(* IEC 61131-3 sources: REFUSR/GP/Refusr.jl/samples (part 18) *)

(* ---- 5-MUX_vitae-roger-ships.st ---- *)
(*
This code implements a shuffled multiplexer with 5 control bits.
The control bits are: Data[N21], Data[N4], Data[N1], Data[N2], Data[N3]
The input bits are: Data[N7], Data[N8], Data[N5], Data[N20], Data[N23], Data[N24], Data[N9], Data[N25], Data[N22], Data[N6], Data[N10], Data[N26], Data[N14], Data[N11], Data[N29], Data[N15], Data[N12], Data[N13], Data[N19], Data[N16], Data[N17], Data[N18], Data[N32], Data[N27], Data[N30], Data[N33], Data[N31], Data[N34], Data[N35], Data[N28], Data[N36], Data[N37]

The symbolic expression is:
((((((((((((((((((((((((((((((((!(((((!(IN21)) & (!(IN4))) & (!(IN1))) & (!(IN2))) & (!(IN3)))) | IN7) & ((!((((IN21 & (!(IN4))) & (!(IN1))) & (!(IN2))) & (!(IN3)))) | IN8)) & ((!(((((!(IN21)) & IN4) & (!(IN1))) & (!(IN2))) & (!(IN3)))) | IN5)) & ((!((((IN21 & IN4) & (!(IN1))) & (!(IN2))) & (!(IN3)))) | IN20)) & ((!(((((!(IN21)) & (!(IN4))) & IN1) & (!(IN2))) & (!(IN3)))) | IN23)) & ((!((((IN21 & (!(IN4))) & IN1) & (!(IN2))) & (!(IN3)))) | IN24)) & ((!(((((!(IN21)) & IN4) & IN1) & (!(IN2))) & (!(IN3)))) | IN9)) & ((!((((IN21 & IN4) & IN1) & (!(IN2))) & (!(IN3)))) | IN25)) & ((!(((((!(IN21)) & (!(IN4))) & (!(IN1))) & IN2) & (!(IN3)))) | IN22)) & ((!((((IN21 & (!(IN4))) & (!(IN1))) & IN2) & (!(IN3)))) | IN6)) & ((!(((((!(IN21)) & IN4) & (!(IN1))) & IN2) & (!(IN3)))) | IN10)) & ((!((((IN21 & IN4) & (!(IN1))) & IN2) & (!(IN3)))) | IN26)) & ((!(((((!(IN21)) & (!(IN4))) & IN1) & IN2) & (!(IN3)))) | IN14)) & ((!((((IN21 & (!(IN4))) & IN1) & IN2) & (!(IN3)))) | IN11)) & ((!(((((!(IN21)) & IN4) & IN1) & IN2) & (!(IN3)))) | IN29)) & ((!((((IN21 & IN4) & IN1) & IN2) & (!(IN3)))) | IN15)) & ((!(((((!(IN21)) & (!(IN4))) & (!(IN1))) & (!(IN2))) & IN3)) | IN12)) & ((!((((IN21 & (!(IN4))) & (!(IN1))) & (!(IN2))) & IN3)) | IN13)) & ((!(((((!(IN21)) & IN4) & (!(IN1))) & (!(IN2))) & IN3)) | IN19)) & ((!((((IN21 & IN4) & (!(IN1))) & (!(IN2))) & IN3)) | IN16)) & ((!(((((!(IN21)) & (!(IN4))) & IN1) & (!(IN2))) & IN3)) | IN17)) & ((!((((IN21 & (!(IN4))) & IN1) & (!(IN2))) & IN3)) | IN18)) & ((!(((((!(IN21)) & IN4) & IN1) & (!(IN2))) & IN3)) | IN32)) & ((!((((IN21 & IN4) & IN1) & (!(IN2))) & IN3)) | IN27)) & ((!(((((!(IN21)) & (!(IN4))) & (!(IN1))) & IN2) & IN3)) | IN30)) & ((!((((IN21 & (!(IN4))) & (!(IN1))) & IN2) & IN3)) | IN33)) & ((!(((((!(IN21)) & IN4) & (!(IN1))) & IN2) & IN3)) | IN31)) & ((!((((IN21 & IN4) & (!(IN1))) & IN2) & IN3)) | IN34)) & ((!(((((!(IN21)) & (!(IN4))) & IN1) & IN2) & IN3)) | IN35)) & ((!((((IN21 & (!(IN4))) & IN1) & IN2) & IN3)) | IN28)) & ((!(((((!(IN21)) & IN4) & IN1) & IN2) & IN3)) | IN36)) & ((!((((IN21 & IN4) & IN1) & IN2) & IN3)) | IN37)

*)

FUNCTION_BLOCK F_CollectInput
  VAR_IN_OUT
      Data : ARRAY[1..40] OF BOOL;
  END_VAR
  VAR_INPUT
      TICK  : BOOL := 0;
      IN1   : BOOL := 0;
      IN2   : BOOL := 0;
      IN3   : BOOL := 0;
      IN4   : BOOL := 0;
      IN5   : BOOL := 0;
      RESET : BOOL := FALSE;
  END_VAR
  VAR_OUTPUT
      Finished : BOOL;
  END_VAR
  VAR
      j    : USINT := 1;
      tock : BOOL  := 0;
  END_VAR
  IF NOT RESET AND tock = NOT TICK THEN
      Data[j]   := IN1;
      Data[j+1] := IN2;
      Data[j+2] := IN3;
      Data[j+3] := IN4;
      Data[j+4] := IN5;
      j := j + 5;
      tock := TICK;
  ELSE
      j := 1;
      tock := 0;
  END_IF;
  Finished := (j > 40);
END_FUNCTION_BLOCK

PROGRAM Boiler
  VAR
    Data  : ARRAY[1..40] OF BOOL;
    Ready : BOOL;
    CollectInput : F_CollectInput;
  END_VAR
  VAR
    TICK     AT %IX1.0 : BOOL;
    IN1      AT %IX0.3 : BOOL;
    IN2      AT %IX0.4 : BOOL;
    IN3      AT %IX0.5 : BOOL;
    IN4      AT %IX0.6 : BOOL;
    IN5      AT %IX0.7 : BOOL;
    OutReady AT %QX0.0 : BOOL := FALSE;
    FeedNext AT %QX0.1 : BOOL := FALSE;
    Out      AT %QX0.2 : BOOL;
  END_VAR
  CollectInput(TICK:=TICK, IN1:=IN1, IN2:=IN2, IN3:=IN3, IN4:=IN4, IN5:=IN5);
  Ready := CollectInput.Finished;
  FeedNext := 1;
  IF Ready THEN
    Out := (((((((((((((((((((((((((((((((((NOT (((((NOT Data[21]) AND (NOT Data[4])) AND (NOT Data[1])) AND (NOT Data[2])) AND (NOT Data[3]))) OR Data[7]) AND ((NOT ((((Data[21] AND (NOT Data[4])) AND (NOT Data[1])) AND (NOT Data[2])) AND (NOT Data[3]))) OR Data[8])) AND ((NOT (((((NOT Data[21]) AND Data[4]) AND (NOT Data[1])) AND (NOT Data[2])) AND (NOT Data[3]))) OR Data[5])) AND ((NOT ((((Data[21] AND Data[4]) AND (NOT Data[1])) AND (NOT Data[2])) AND (NOT Data[3]))) OR Data[20])) AND ((NOT (((((NOT Data[21]) AND (NOT Data[4])) AND Data[1]) AND (NOT Data[2])) AND (NOT Data[3]))) OR Data[23])) AND ((NOT ((((Data[21] AND (NOT Data[4])) AND Data[1]) AND (NOT Data[2])) AND (NOT Data[3]))) OR Data[24])) AND ((NOT (((((NOT Data[21]) AND Data[4]) AND Data[1]) AND (NOT Data[2])) AND (NOT Data[3]))) OR Data[9])) AND ((NOT ((((Data[21] AND Data[4]) AND Data[1]) AND (NOT Data[2])) AND (NOT Data[3]))) OR Data[25])) AND ((NOT (((((NOT Data[21]) AND (NOT Data[4])) AND (NOT Data[1])) AND Data[2]) AND (NOT Data[3]))) OR Data[22])) AND ((NOT ((((Data[21] AND (NOT Data[4])) AND (NOT Data[1])) AND Data[2]) AND (NOT Data[3]))) OR Data[6])) AND ((NOT (((((NOT Data[21]) AND Data[4]) AND (NOT Data[1])) AND Data[2]) AND (NOT Data[3]))) OR Data[10])) AND ((NOT ((((Data[21] AND Data[4]) AND (NOT Data[1])) AND Data[2]) AND (NOT Data[3]))) OR Data[26])) AND ((NOT (((((NOT Data[21]) AND (NOT Data[4])) AND Data[1]) AND Data[2]) AND (NOT Data[3]))) OR Data[14])) AND ((NOT ((((Data[21] AND (NOT Data[4])) AND Data[1]) AND Data[2]) AND (NOT Data[3]))) OR Data[11])) AND ((NOT (((((NOT Data[21]) AND Data[4]) AND Data[1]) AND Data[2]) AND (NOT Data[3]))) OR Data[29])) AND ((NOT ((((Data[21] AND Data[4]) AND Data[1]) AND Data[2]) AND (NOT Data[3]))) OR Data[15])) AND ((NOT (((((NOT Data[21]) AND (NOT Data[4])) AND (NOT Data[1])) AND (NOT Data[2])) AND Data[3])) OR Data[12])) AND ((NOT ((((Data[21] AND (NOT Data[4])) AND (NOT Data[1])) AND (NOT Data[2])) AND Data[3])) OR Data[13])) AND ((NOT (((((NOT Data[21]) AND Data[4]) AND (NOT Data[1])) AND (NOT Data[2])) AND Data[3])) OR Data[19])) AND ((NOT ((((Data[21] AND Data[4]) AND (NOT Data[1])) AND (NOT Data[2])) AND Data[3])) OR Data[16])) AND ((NOT (((((NOT Data[21]) AND (NOT Data[4])) AND Data[1]) AND (NOT Data[2])) AND Data[3])) OR Data[17])) AND ((NOT ((((Data[21] AND (NOT Data[4])) AND Data[1]) AND (NOT Data[2])) AND Data[3])) OR Data[18])) AND ((NOT (((((NOT Data[21]) AND Data[4]) AND Data[1]) AND (NOT Data[2])) AND Data[3])) OR Data[32])) AND ((NOT ((((Data[21] AND Data[4]) AND Data[1]) AND (NOT Data[2])) AND Data[3])) OR Data[27])) AND ((NOT (((((NOT Data[21]) AND (NOT Data[4])) AND (NOT Data[1])) AND Data[2]) AND Data[3])) OR Data[30])) AND ((NOT ((((Data[21] AND (NOT Data[4])) AND (NOT Data[1])) AND Data[2]) AND Data[3])) OR Data[33])) AND ((NOT (((((NOT Data[21]) AND Data[4]) AND (NOT Data[1])) AND Data[2]) AND Data[3])) OR Data[31])) AND ((NOT ((((Data[21] AND Data[4]) AND (NOT Data[1])) AND Data[2]) AND Data[3])) OR Data[34])) AND ((NOT (((((NOT Data[21]) AND (NOT Data[4])) AND Data[1]) AND Data[2]) AND Data[3])) OR Data[35])) AND ((NOT ((((Data[21] AND (NOT Data[4])) AND Data[1]) AND Data[2]) AND Data[3])) OR Data[28])) AND ((NOT (((((NOT Data[21]) AND Data[4]) AND Data[1]) AND Data[2]) AND Data[3])) OR Data[36])) AND ((NOT ((((Data[21] AND Data[4]) AND Data[1]) AND Data[2]) AND Data[3])) OR Data[37]));
    OutReady := 1;
    CollectInput(RESET:=TRUE);
  END_IF;
END_PROGRAM

CONFIGURATION Config0
  RESOURCE Res0 ON PLC
    TASK task0(INTERVAL := T#20ms,PRIORITY := 0);
    PROGRAM instance0 WITH task0 : Boiler;
  END_RESOURCE
END_CONFIGURATION

(* ---- 5-MUX_vodka-chive-wrier.st ---- *)
(*
This code implements a shuffled multiplexer with 5 control bits.
The control bits are: Data[N2], Data[N1], Data[N23], Data[N3], Data[N20]
The input bits are: Data[N6], Data[N11], Data[N7], Data[N5], Data[N22], Data[N21], Data[N24], Data[N25], Data[N8], Data[N4], Data[N9], Data[N10], Data[N12], Data[N13], Data[N26], Data[N27], Data[N28], Data[N15], Data[N29], Data[N14], Data[N18], Data[N34], Data[N31], Data[N16], Data[N17], Data[N19], Data[N35], Data[N32], Data[N30], Data[N37], Data[N36], Data[N33]

The symbolic expression is:
((((((((((((((((((((((((((((((((!(((((!(IN2)) & (!(IN1))) & (!(IN23))) & (!(IN3))) & (!(IN20)))) | IN6) & ((!((((IN2 & (!(IN1))) & (!(IN23))) & (!(IN3))) & (!(IN20)))) | IN11)) & ((!(((((!(IN2)) & IN1) & (!(IN23))) & (!(IN3))) & (!(IN20)))) | IN7)) & ((!((((IN2 & IN1) & (!(IN23))) & (!(IN3))) & (!(IN20)))) | IN5)) & ((!(((((!(IN2)) & (!(IN1))) & IN23) & (!(IN3))) & (!(IN20)))) | IN22)) & ((!((((IN2 & (!(IN1))) & IN23) & (!(IN3))) & (!(IN20)))) | IN21)) & ((!(((((!(IN2)) & IN1) & IN23) & (!(IN3))) & (!(IN20)))) | IN24)) & ((!((((IN2 & IN1) & IN23) & (!(IN3))) & (!(IN20)))) | IN25)) & ((!(((((!(IN2)) & (!(IN1))) & (!(IN23))) & IN3) & (!(IN20)))) | IN8)) & ((!((((IN2 & (!(IN1))) & (!(IN23))) & IN3) & (!(IN20)))) | IN4)) & ((!(((((!(IN2)) & IN1) & (!(IN23))) & IN3) & (!(IN20)))) | IN9)) & ((!((((IN2 & IN1) & (!(IN23))) & IN3) & (!(IN20)))) | IN10)) & ((!(((((!(IN2)) & (!(IN1))) & IN23) & IN3) & (!(IN20)))) | IN12)) & ((!((((IN2 & (!(IN1))) & IN23) & IN3) & (!(IN20)))) | IN13)) & ((!(((((!(IN2)) & IN1) & IN23) & IN3) & (!(IN20)))) | IN26)) & ((!((((IN2 & IN1) & IN23) & IN3) & (!(IN20)))) | IN27)) & ((!(((((!(IN2)) & (!(IN1))) & (!(IN23))) & (!(IN3))) & IN20)) | IN28)) & ((!((((IN2 & (!(IN1))) & (!(IN23))) & (!(IN3))) & IN20)) | IN15)) & ((!(((((!(IN2)) & IN1) & (!(IN23))) & (!(IN3))) & IN20)) | IN29)) & ((!((((IN2 & IN1) & (!(IN23))) & (!(IN3))) & IN20)) | IN14)) & ((!(((((!(IN2)) & (!(IN1))) & IN23) & (!(IN3))) & IN20)) | IN18)) & ((!((((IN2 & (!(IN1))) & IN23) & (!(IN3))) & IN20)) | IN34)) & ((!(((((!(IN2)) & IN1) & IN23) & (!(IN3))) & IN20)) | IN31)) & ((!((((IN2 & IN1) & IN23) & (!(IN3))) & IN20)) | IN16)) & ((!(((((!(IN2)) & (!(IN1))) & (!(IN23))) & IN3) & IN20)) | IN17)) & ((!((((IN2 & (!(IN1))) & (!(IN23))) & IN3) & IN20)) | IN19)) & ((!(((((!(IN2)) & IN1) & (!(IN23))) & IN3) & IN20)) | IN35)) & ((!((((IN2 & IN1) & (!(IN23))) & IN3) & IN20)) | IN32)) & ((!(((((!(IN2)) & (!(IN1))) & IN23) & IN3) & IN20)) | IN30)) & ((!((((IN2 & (!(IN1))) & IN23) & IN3) & IN20)) | IN37)) & ((!(((((!(IN2)) & IN1) & IN23) & IN3) & IN20)) | IN36)) & ((!((((IN2 & IN1) & IN23) & IN3) & IN20)) | IN33)

*)

FUNCTION_BLOCK F_CollectInput
  VAR_IN_OUT
      Data : ARRAY[1..40] OF BOOL;
  END_VAR
  VAR_INPUT
      TICK  : BOOL := 0;
      IN1   : BOOL := 0;
      IN2   : BOOL := 0;
      IN3   : BOOL := 0;
      IN4   : BOOL := 0;
      IN5   : BOOL := 0;
      RESET : BOOL := FALSE;
  END_VAR
  VAR_OUTPUT
      Finished : BOOL;
  END_VAR
  VAR
      j    : USINT := 1;
      tock : BOOL  := 0;
  END_VAR
  IF NOT RESET AND tock = NOT TICK THEN
      Data[j]   := IN1;
      Data[j+1] := IN2;
      Data[j+2] := IN3;
      Data[j+3] := IN4;
      Data[j+4] := IN5;
      j := j + 5;
      tock := TICK;
  ELSE
      j := 1;
      tock := 0;
  END_IF;
  Finished := (j > 40);
END_FUNCTION_BLOCK

PROGRAM Boiler
  VAR
    Data  : ARRAY[1..40] OF BOOL;
    Ready : BOOL;
    CollectInput : F_CollectInput;
  END_VAR
  VAR
    TICK     AT %IX1.0 : BOOL;
    IN1      AT %IX0.3 : BOOL;
    IN2      AT %IX0.4 : BOOL;
    IN3      AT %IX0.5 : BOOL;
    IN4      AT %IX0.6 : BOOL;
    IN5      AT %IX0.7 : BOOL;
    OutReady AT %QX0.0 : BOOL := FALSE;
    FeedNext AT %QX0.1 : BOOL := FALSE;
    Out      AT %QX0.2 : BOOL;
  END_VAR
  CollectInput(TICK:=TICK, IN1:=IN1, IN2:=IN2, IN3:=IN3, IN4:=IN4, IN5:=IN5);
  Ready := CollectInput.Finished;
  FeedNext := 1;
  IF Ready THEN
    Out := (((((((((((((((((((((((((((((((((NOT (((((NOT Data[2]) AND (NOT Data[1])) AND (NOT Data[23])) AND (NOT Data[3])) AND (NOT Data[20]))) OR Data[6]) AND ((NOT ((((Data[2] AND (NOT Data[1])) AND (NOT Data[23])) AND (NOT Data[3])) AND (NOT Data[20]))) OR Data[11])) AND ((NOT (((((NOT Data[2]) AND Data[1]) AND (NOT Data[23])) AND (NOT Data[3])) AND (NOT Data[20]))) OR Data[7])) AND ((NOT ((((Data[2] AND Data[1]) AND (NOT Data[23])) AND (NOT Data[3])) AND (NOT Data[20]))) OR Data[5])) AND ((NOT (((((NOT Data[2]) AND (NOT Data[1])) AND Data[23]) AND (NOT Data[3])) AND (NOT Data[20]))) OR Data[22])) AND ((NOT ((((Data[2] AND (NOT Data[1])) AND Data[23]) AND (NOT Data[3])) AND (NOT Data[20]))) OR Data[21])) AND ((NOT (((((NOT Data[2]) AND Data[1]) AND Data[23]) AND (NOT Data[3])) AND (NOT Data[20]))) OR Data[24])) AND ((NOT ((((Data[2] AND Data[1]) AND Data[23]) AND (NOT Data[3])) AND (NOT Data[20]))) OR Data[25])) AND ((NOT (((((NOT Data[2]) AND (NOT Data[1])) AND (NOT Data[23])) AND Data[3]) AND (NOT Data[20]))) OR Data[8])) AND ((NOT ((((Data[2] AND (NOT Data[1])) AND (NOT Data[23])) AND Data[3]) AND (NOT Data[20]))) OR Data[4])) AND ((NOT (((((NOT Data[2]) AND Data[1]) AND (NOT Data[23])) AND Data[3]) AND (NOT Data[20]))) OR Data[9])) AND ((NOT ((((Data[2] AND Data[1]) AND (NOT Data[23])) AND Data[3]) AND (NOT Data[20]))) OR Data[10])) AND ((NOT (((((NOT Data[2]) AND (NOT Data[1])) AND Data[23]) AND Data[3]) AND (NOT Data[20]))) OR Data[12])) AND ((NOT ((((Data[2] AND (NOT Data[1])) AND Data[23]) AND Data[3]) AND (NOT Data[20]))) OR Data[13])) AND ((NOT (((((NOT Data[2]) AND Data[1]) AND Data[23]) AND Data[3]) AND (NOT Data[20]))) OR Data[26])) AND ((NOT ((((Data[2] AND Data[1]) AND Data[23]) AND Data[3]) AND (NOT Data[20]))) OR Data[27])) AND ((NOT (((((NOT Data[2]) AND (NOT Data[1])) AND (NOT Data[23])) AND (NOT Data[3])) AND Data[20])) OR Data[28])) AND ((NOT ((((Data[2] AND (NOT Data[1])) AND (NOT Data[23])) AND (NOT Data[3])) AND Data[20])) OR Data[15])) AND ((NOT (((((NOT Data[2]) AND Data[1]) AND (NOT Data[23])) AND (NOT Data[3])) AND Data[20])) OR Data[29])) AND ((NOT ((((Data[2] AND Data[1]) AND (NOT Data[23])) AND (NOT Data[3])) AND Data[20])) OR Data[14])) AND ((NOT (((((NOT Data[2]) AND (NOT Data[1])) AND Data[23]) AND (NOT Data[3])) AND Data[20])) OR Data[18])) AND ((NOT ((((Data[2] AND (NOT Data[1])) AND Data[23]) AND (NOT Data[3])) AND Data[20])) OR Data[34])) AND ((NOT (((((NOT Data[2]) AND Data[1]) AND Data[23]) AND (NOT Data[3])) AND Data[20])) OR Data[31])) AND ((NOT ((((Data[2] AND Data[1]) AND Data[23]) AND (NOT Data[3])) AND Data[20])) OR Data[16])) AND ((NOT (((((NOT Data[2]) AND (NOT Data[1])) AND (NOT Data[23])) AND Data[3]) AND Data[20])) OR Data[17])) AND ((NOT ((((Data[2] AND (NOT Data[1])) AND (NOT Data[23])) AND Data[3]) AND Data[20])) OR Data[19])) AND ((NOT (((((NOT Data[2]) AND Data[1]) AND (NOT Data[23])) AND Data[3]) AND Data[20])) OR Data[35])) AND ((NOT ((((Data[2] AND Data[1]) AND (NOT Data[23])) AND Data[3]) AND Data[20])) OR Data[32])) AND ((NOT (((((NOT Data[2]) AND (NOT Data[1])) AND Data[23]) AND Data[3]) AND Data[20])) OR Data[30])) AND ((NOT ((((Data[2] AND (NOT Data[1])) AND Data[23]) AND Data[3]) AND Data[20])) OR Data[37])) AND ((NOT (((((NOT Data[2]) AND Data[1]) AND Data[23]) AND Data[3]) AND Data[20])) OR Data[36])) AND ((NOT ((((Data[2] AND Data[1]) AND Data[23]) AND Data[3]) AND Data[20])) OR Data[33]));
    OutReady := 1;
    CollectInput(RESET:=TRUE);
  END_IF;
END_PROGRAM

CONFIGURATION Config0
  RESOURCE Res0 ON PLC
    TASK task0(INTERVAL := T#20ms,PRIORITY := 0);
    PROGRAM instance0 WITH task0 : Boiler;
  END_RESOURCE
END_CONFIGURATION

(* ---- 5-MUX_wager-river-honky.st ---- *)
(*
This code implements a shuffled multiplexer with 5 control bits.
The control bits are: Data[N22], Data[N21], Data[N2], Data[N20], Data[N5]
The input bits are: Data[N3], Data[N6], Data[N4], Data[N8], Data[N23], Data[N9], Data[N7], Data[N24], Data[N25], Data[N1], Data[N14], Data[N26], Data[N28], Data[N15], Data[N13], Data[N27], Data[N10], Data[N29], Data[N17], Data[N33], Data[N11], Data[N12], Data[N16], Data[N30], Data[N19], Data[N18], Data[N31], Data[N36], Data[N37], Data[N34], Data[N32], Data[N35]

The symbolic expression is:
((((((((((((((((((((((((((((((((!(((((!(IN22)) & (!(IN21))) & (!(IN2))) & (!(IN20))) & (!(IN5)))) | IN3) & ((!((((IN22 & (!(IN21))) & (!(IN2))) & (!(IN20))) & (!(IN5)))) | IN6)) & ((!(((((!(IN22)) & IN21) & (!(IN2))) & (!(IN20))) & (!(IN5)))) | IN4)) & ((!((((IN22 & IN21) & (!(IN2))) & (!(IN20))) & (!(IN5)))) | IN8)) & ((!(((((!(IN22)) & (!(IN21))) & IN2) & (!(IN20))) & (!(IN5)))) | IN23)) & ((!((((IN22 & (!(IN21))) & IN2) & (!(IN20))) & (!(IN5)))) | IN9)) & ((!(((((!(IN22)) & IN21) & IN2) & (!(IN20))) & (!(IN5)))) | IN7)) & ((!((((IN22 & IN21) & IN2) & (!(IN20))) & (!(IN5)))) | IN24)) & ((!(((((!(IN22)) & (!(IN21))) & (!(IN2))) & IN20) & (!(IN5)))) | IN25)) & ((!((((IN22 & (!(IN21))) & (!(IN2))) & IN20) & (!(IN5)))) | IN1)) & ((!(((((!(IN22)) & IN21) & (!(IN2))) & IN20) & (!(IN5)))) | IN14)) & ((!((((IN22 & IN21) & (!(IN2))) & IN20) & (!(IN5)))) | IN26)) & ((!(((((!(IN22)) & (!(IN21))) & IN2) & IN20) & (!(IN5)))) | IN28)) & ((!((((IN22 & (!(IN21))) & IN2) & IN20) & (!(IN5)))) | IN15)) & ((!(((((!(IN22)) & IN21) & IN2) & IN20) & (!(IN5)))) | IN13)) & ((!((((IN22 & IN21) & IN2) & IN20) & (!(IN5)))) | IN27)) & ((!(((((!(IN22)) & (!(IN21))) & (!(IN2))) & (!(IN20))) & IN5)) | IN10)) & ((!((((IN22 & (!(IN21))) & (!(IN2))) & (!(IN20))) & IN5)) | IN29)) & ((!(((((!(IN22)) & IN21) & (!(IN2))) & (!(IN20))) & IN5)) | IN17)) & ((!((((IN22 & IN21) & (!(IN2))) & (!(IN20))) & IN5)) | IN33)) & ((!(((((!(IN22)) & (!(IN21))) & IN2) & (!(IN20))) & IN5)) | IN11)) & ((!((((IN22 & (!(IN21))) & IN2) & (!(IN20))) & IN5)) | IN12)) & ((!(((((!(IN22)) & IN21) & IN2) & (!(IN20))) & IN5)) | IN16)) & ((!((((IN22 & IN21) & IN2) & (!(IN20))) & IN5)) | IN30)) & ((!(((((!(IN22)) & (!(IN21))) & (!(IN2))) & IN20) & IN5)) | IN19)) & ((!((((IN22 & (!(IN21))) & (!(IN2))) & IN20) & IN5)) | IN18)) & ((!(((((!(IN22)) & IN21) & (!(IN2))) & IN20) & IN5)) | IN31)) & ((!((((IN22 & IN21) & (!(IN2))) & IN20) & IN5)) | IN36)) & ((!(((((!(IN22)) & (!(IN21))) & IN2) & IN20) & IN5)) | IN37)) & ((!((((IN22 & (!(IN21))) & IN2) & IN20) & IN5)) | IN34)) & ((!(((((!(IN22)) & IN21) & IN2) & IN20) & IN5)) | IN32)) & ((!((((IN22 & IN21) & IN2) & IN20) & IN5)) | IN35)

*)

FUNCTION_BLOCK F_CollectInput
  VAR_IN_OUT
      Data : ARRAY[1..40] OF BOOL;
  END_VAR
  VAR_INPUT
      TICK  : BOOL := 0;
      IN1   : BOOL := 0;
      IN2   : BOOL := 0;
      IN3   : BOOL := 0;
      IN4   : BOOL := 0;
      IN5   : BOOL := 0;
      RESET : BOOL := FALSE;
  END_VAR
  VAR_OUTPUT
      Finished : BOOL;
  END_VAR
  VAR
      j    : USINT := 1;
      tock : BOOL  := 0;
  END_VAR
  IF NOT RESET AND tock = NOT TICK THEN
      Data[j]   := IN1;
      Data[j+1] := IN2;
      Data[j+2] := IN3;
      Data[j+3] := IN4;
      Data[j+4] := IN5;
      j := j + 5;
      tock := TICK;
  ELSE
      j := 1;
      tock := 0;
  END_IF;
  Finished := (j > 40);
END_FUNCTION_BLOCK

PROGRAM Boiler
  VAR
    Data  : ARRAY[1..40] OF BOOL;
    Ready : BOOL;
    CollectInput : F_CollectInput;
  END_VAR
  VAR
    TICK     AT %IX1.0 : BOOL;
    IN1      AT %IX0.3 : BOOL;
    IN2      AT %IX0.4 : BOOL;
    IN3      AT %IX0.5 : BOOL;
    IN4      AT %IX0.6 : BOOL;
    IN5      AT %IX0.7 : BOOL;
    OutReady AT %QX0.0 : BOOL := FALSE;
    FeedNext AT %QX0.1 : BOOL := FALSE;
    Out      AT %QX0.2 : BOOL;
  END_VAR
  CollectInput(TICK:=TICK, IN1:=IN1, IN2:=IN2, IN3:=IN3, IN4:=IN4, IN5:=IN5);
  Ready := CollectInput.Finished;
  FeedNext := 1;
  IF Ready THEN
    Out := (((((((((((((((((((((((((((((((((NOT (((((NOT Data[22]) AND (NOT Data[21])) AND (NOT Data[2])) AND (NOT Data[20])) AND (NOT Data[5]))) OR Data[3]) AND ((NOT ((((Data[22] AND (NOT Data[21])) AND (NOT Data[2])) AND (NOT Data[20])) AND (NOT Data[5]))) OR Data[6])) AND ((NOT (((((NOT Data[22]) AND Data[21]) AND (NOT Data[2])) AND (NOT Data[20])) AND (NOT Data[5]))) OR Data[4])) AND ((NOT ((((Data[22] AND Data[21]) AND (NOT Data[2])) AND (NOT Data[20])) AND (NOT Data[5]))) OR Data[8])) AND ((NOT (((((NOT Data[22]) AND (NOT Data[21])) AND Data[2]) AND (NOT Data[20])) AND (NOT Data[5]))) OR Data[23])) AND ((NOT ((((Data[22] AND (NOT Data[21])) AND Data[2]) AND (NOT Data[20])) AND (NOT Data[5]))) OR Data[9])) AND ((NOT (((((NOT Data[22]) AND Data[21]) AND Data[2]) AND (NOT Data[20])) AND (NOT Data[5]))) OR Data[7])) AND ((NOT ((((Data[22] AND Data[21]) AND Data[2]) AND (NOT Data[20])) AND (NOT Data[5]))) OR Data[24])) AND ((NOT (((((NOT Data[22]) AND (NOT Data[21])) AND (NOT Data[2])) AND Data[20]) AND (NOT Data[5]))) OR Data[25])) AND ((NOT ((((Data[22] AND (NOT Data[21])) AND (NOT Data[2])) AND Data[20]) AND (NOT Data[5]))) OR Data[1])) AND ((NOT (((((NOT Data[22]) AND Data[21]) AND (NOT Data[2])) AND Data[20]) AND (NOT Data[5]))) OR Data[14])) AND ((NOT ((((Data[22] AND Data[21]) AND (NOT Data[2])) AND Data[20]) AND (NOT Data[5]))) OR Data[26])) AND ((NOT (((((NOT Data[22]) AND (NOT Data[21])) AND Data[2]) AND Data[20]) AND (NOT Data[5]))) OR Data[28])) AND ((NOT ((((Data[22] AND (NOT Data[21])) AND Data[2]) AND Data[20]) AND (NOT Data[5]))) OR Data[15])) AND ((NOT (((((NOT Data[22]) AND Data[21]) AND Data[2]) AND Data[20]) AND (NOT Data[5]))) OR Data[13])) AND ((NOT ((((Data[22] AND Data[21]) AND Data[2]) AND Data[20]) AND (NOT Data[5]))) OR Data[27])) AND ((NOT (((((NOT Data[22]) AND (NOT Data[21])) AND (NOT Data[2])) AND (NOT Data[20])) AND Data[5])) OR Data[10])) AND ((NOT ((((Data[22] AND (NOT Data[21])) AND (NOT Data[2])) AND (NOT Data[20])) AND Data[5])) OR Data[29])) AND ((NOT (((((NOT Data[22]) AND Data[21]) AND (NOT Data[2])) AND (NOT Data[20])) AND Data[5])) OR Data[17])) AND ((NOT ((((Data[22] AND Data[21]) AND (NOT Data[2])) AND (NOT Data[20])) AND Data[5])) OR Data[33])) AND ((NOT (((((NOT Data[22]) AND (NOT Data[21])) AND Data[2]) AND (NOT Data[20])) AND Data[5])) OR Data[11])) AND ((NOT ((((Data[22] AND (NOT Data[21])) AND Data[2]) AND (NOT Data[20])) AND Data[5])) OR Data[12])) AND ((NOT (((((NOT Data[22]) AND Data[21]) AND Data[2]) AND (NOT Data[20])) AND Data[5])) OR Data[16])) AND ((NOT ((((Data[22] AND Data[21]) AND Data[2]) AND (NOT Data[20])) AND Data[5])) OR Data[30])) AND ((NOT (((((NOT Data[22]) AND (NOT Data[21])) AND (NOT Data[2])) AND Data[20]) AND Data[5])) OR Data[19])) AND ((NOT ((((Data[22] AND (NOT Data[21])) AND (NOT Data[2])) AND Data[20]) AND Data[5])) OR Data[18])) AND ((NOT (((((NOT Data[22]) AND Data[21]) AND (NOT Data[2])) AND Data[20]) AND Data[5])) OR Data[31])) AND ((NOT ((((Data[22] AND Data[21]) AND (NOT Data[2])) AND Data[20]) AND Data[5])) OR Data[36])) AND ((NOT (((((NOT Data[22]) AND (NOT Data[21])) AND Data[2]) AND Data[20]) AND Data[5])) OR Data[37])) AND ((NOT ((((Data[22] AND (NOT Data[21])) AND Data[2]) AND Data[20]) AND Data[5])) OR Data[34])) AND ((NOT (((((NOT Data[22]) AND Data[21]) AND Data[2]) AND Data[20]) AND Data[5])) OR Data[32])) AND ((NOT ((((Data[22] AND Data[21]) AND Data[2]) AND Data[20]) AND Data[5])) OR Data[35]));
    OutReady := 1;
    CollectInput(RESET:=TRUE);
  END_IF;
END_PROGRAM

CONFIGURATION Config0
  RESOURCE Res0 ON PLC
    TASK task0(INTERVAL := T#20ms,PRIORITY := 0);
    PROGRAM instance0 WITH task0 : Boiler;
  END_RESOURCE
END_CONFIGURATION

(* ---- 5-MUX_waken-moldy-alway.st ---- *)
(*
This code implements a shuffled multiplexer with 5 control bits.
The control bits are: Data[N1], Data[N2], Data[N3], Data[N4], Data[N23]
The input bits are: Data[N22], Data[N21], Data[N5], Data[N12], Data[N6], Data[N9], Data[N7], Data[N20], Data[N14], Data[N25], Data[N11], Data[N24], Data[N16], Data[N26], Data[N13], Data[N27], Data[N15], Data[N8], Data[N17], Data[N10], Data[N18], Data[N28], Data[N19], Data[N29], Data[N30], Data[N31], Data[N32], Data[N33], Data[N34], Data[N35], Data[N36], Data[N37]

The symbolic expression is:
((((((((((((((((((((((((((((((((!(((((!(IN1)) & (!(IN2))) & (!(IN3))) & (!(IN4))) & (!(IN23)))) | IN22) & ((!((((IN1 & (!(IN2))) & (!(IN3))) & (!(IN4))) & (!(IN23)))) | IN21)) & ((!(((((!(IN1)) & IN2) & (!(IN3))) & (!(IN4))) & (!(IN23)))) | IN5)) & ((!((((IN1 & IN2) & (!(IN3))) & (!(IN4))) & (!(IN23)))) | IN12)) & ((!(((((!(IN1)) & (!(IN2))) & IN3) & (!(IN4))) & (!(IN23)))) | IN6)) & ((!((((IN1 & (!(IN2))) & IN3) & (!(IN4))) & (!(IN23)))) | IN9)) & ((!(((((!(IN1)) & IN2) & IN3) & (!(IN4))) & (!(IN23)))) | IN7)) & ((!((((IN1 & IN2) & IN3) & (!(IN4))) & (!(IN23)))) | IN20)) & ((!(((((!(IN1)) & (!(IN2))) & (!(IN3))) & IN4) & (!(IN23)))) | IN14)) & ((!((((IN1 & (!(IN2))) & (!(IN3))) & IN4) & (!(IN23)))) | IN25)) & ((!(((((!(IN1)) & IN2) & (!(IN3))) & IN4) & (!(IN23)))) | IN11)) & ((!((((IN1 & IN2) & (!(IN3))) & IN4) & (!(IN23)))) | IN24)) & ((!(((((!(IN1)) & (!(IN2))) & IN3) & IN4) & (!(IN23)))) | IN16)) & ((!((((IN1 & (!(IN2))) & IN3) & IN4) & (!(IN23)))) | IN26)) & ((!(((((!(IN1)) & IN2) & IN3) & IN4) & (!(IN23)))) | IN13)) & ((!((((IN1 & IN2) & IN3) & IN4) & (!(IN23)))) | IN27)) & ((!(((((!(IN1)) & (!(IN2))) & (!(IN3))) & (!(IN4))) & IN23)) | IN15)) & ((!((((IN1 & (!(IN2))) & (!(IN3))) & (!(IN4))) & IN23)) | IN8)) & ((!(((((!(IN1)) & IN2) & (!(IN3))) & (!(IN4))) & IN23)) | IN17)) & ((!((((IN1 & IN2) & (!(IN3))) & (!(IN4))) & IN23)) | IN10)) & ((!(((((!(IN1)) & (!(IN2))) & IN3) & (!(IN4))) & IN23)) | IN18)) & ((!((((IN1 & (!(IN2))) & IN3) & (!(IN4))) & IN23)) | IN28)) & ((!(((((!(IN1)) & IN2) & IN3) & (!(IN4))) & IN23)) | IN19)) & ((!((((IN1 & IN2) & IN3) & (!(IN4))) & IN23)) | IN29)) & ((!(((((!(IN1)) & (!(IN2))) & (!(IN3))) & IN4) & IN23)) | IN30)) & ((!((((IN1 & (!(IN2))) & (!(IN3))) & IN4) & IN23)) | IN31)) & ((!(((((!(IN1)) & IN2) & (!(IN3))) & IN4) & IN23)) | IN32)) & ((!((((IN1 & IN2) & (!(IN3))) & IN4) & IN23)) | IN33)) & ((!(((((!(IN1)) & (!(IN2))) & IN3) & IN4) & IN23)) | IN34)) & ((!((((IN1 & (!(IN2))) & IN3) & IN4) & IN23)) | IN35)) & ((!(((((!(IN1)) & IN2) & IN3) & IN4) & IN23)) | IN36)) & ((!((((IN1 & IN2) & IN3) & IN4) & IN23)) | IN37)

*)

FUNCTION_BLOCK F_CollectInput
  VAR_IN_OUT
      Data : ARRAY[1..40] OF BOOL;
  END_VAR
  VAR_INPUT
      TICK  : BOOL := 0;
      IN1   : BOOL := 0;
      IN2   : BOOL := 0;
      IN3   : BOOL := 0;
      IN4   : BOOL := 0;
      IN5   : BOOL := 0;
      RESET : BOOL := FALSE;
  END_VAR
  VAR_OUTPUT
      Finished : BOOL;
  END_VAR
  VAR
      j    : USINT := 1;
      tock : BOOL  := 0;
  END_VAR
  IF NOT RESET AND tock = NOT TICK THEN
      Data[j]   := IN1;
      Data[j+1] := IN2;
      Data[j+2] := IN3;
      Data[j+3] := IN4;
      Data[j+4] := IN5;
      j := j + 5;
      tock := TICK;
  ELSE
      j := 1;
      tock := 0;
  END_IF;
  Finished := (j > 40);
END_FUNCTION_BLOCK

PROGRAM Boiler
  VAR
    Data  : ARRAY[1..40] OF BOOL;
    Ready : BOOL;
    CollectInput : F_CollectInput;
  END_VAR
  VAR
    TICK     AT %IX1.0 : BOOL;
    IN1      AT %IX0.3 : BOOL;
    IN2      AT %IX0.4 : BOOL;
    IN3      AT %IX0.5 : BOOL;
    IN4      AT %IX0.6 : BOOL;
    IN5      AT %IX0.7 : BOOL;
    OutReady AT %QX0.0 : BOOL := FALSE;
    FeedNext AT %QX0.1 : BOOL := FALSE;
    Out      AT %QX0.2 : BOOL;
  END_VAR
  CollectInput(TICK:=TICK, IN1:=IN1, IN2:=IN2, IN3:=IN3, IN4:=IN4, IN5:=IN5);
  Ready := CollectInput.Finished;
  FeedNext := 1;
  IF Ready THEN
    Out := (((((((((((((((((((((((((((((((((NOT (((((NOT Data[1]) AND (NOT Data[2])) AND (NOT Data[3])) AND (NOT Data[4])) AND (NOT Data[23]))) OR Data[22]) AND ((NOT ((((Data[1] AND (NOT Data[2])) AND (NOT Data[3])) AND (NOT Data[4])) AND (NOT Data[23]))) OR Data[21])) AND ((NOT (((((NOT Data[1]) AND Data[2]) AND (NOT Data[3])) AND (NOT Data[4])) AND (NOT Data[23]))) OR Data[5])) AND ((NOT ((((Data[1] AND Data[2]) AND (NOT Data[3])) AND (NOT Data[4])) AND (NOT Data[23]))) OR Data[12])) AND ((NOT (((((NOT Data[1]) AND (NOT Data[2])) AND Data[3]) AND (NOT Data[4])) AND (NOT Data[23]))) OR Data[6])) AND ((NOT ((((Data[1] AND (NOT Data[2])) AND Data[3]) AND (NOT Data[4])) AND (NOT Data[23]))) OR Data[9])) AND ((NOT (((((NOT Data[1]) AND Data[2]) AND Data[3]) AND (NOT Data[4])) AND (NOT Data[23]))) OR Data[7])) AND ((NOT ((((Data[1] AND Data[2]) AND Data[3]) AND (NOT Data[4])) AND (NOT Data[23]))) OR Data[20])) AND ((NOT (((((NOT Data[1]) AND (NOT Data[2])) AND (NOT Data[3])) AND Data[4]) AND (NOT Data[23]))) OR Data[14])) AND ((NOT ((((Data[1] AND (NOT Data[2])) AND (NOT Data[3])) AND Data[4]) AND (NOT Data[23]))) OR Data[25])) AND ((NOT (((((NOT Data[1]) AND Data[2]) AND (NOT Data[3])) AND Data[4]) AND (NOT Data[23]))) OR Data[11])) AND ((NOT ((((Data[1] AND Data[2]) AND (NOT Data[3])) AND Data[4]) AND (NOT Data[23]))) OR Data[24])) AND ((NOT (((((NOT Data[1]) AND (NOT Data[2])) AND Data[3]) AND Data[4]) AND (NOT Data[23]))) OR Data[16])) AND ((NOT ((((Data[1] AND (NOT Data[2])) AND Data[3]) AND Data[4]) AND (NOT Data[23]))) OR Data[26])) AND ((NOT (((((NOT Data[1]) AND Data[2]) AND Data[3]) AND Data[4]) AND (NOT Data[23]))) OR Data[13])) AND ((NOT ((((Data[1] AND Data[2]) AND Data[3]) AND Data[4]) AND (NOT Data[23]))) OR Data[27])) AND ((NOT (((((NOT Data[1]) AND (NOT Data[2])) AND (NOT Data[3])) AND (NOT Data[4])) AND Data[23])) OR Data[15])) AND ((NOT ((((Data[1] AND (NOT Data[2])) AND (NOT Data[3])) AND (NOT Data[4])) AND Data[23])) OR Data[8])) AND ((NOT (((((NOT Data[1]) AND Data[2]) AND (NOT Data[3])) AND (NOT Data[4])) AND Data[23])) OR Data[17])) AND ((NOT ((((Data[1] AND Data[2]) AND (NOT Data[3])) AND (NOT Data[4])) AND Data[23])) OR Data[10])) AND ((NOT (((((NOT Data[1]) AND (NOT Data[2])) AND Data[3]) AND (NOT Data[4])) AND Data[23])) OR Data[18])) AND ((NOT ((((Data[1] AND (NOT Data[2])) AND Data[3]) AND (NOT Data[4])) AND Data[23])) OR Data[28])) AND ((NOT (((((NOT Data[1]) AND Data[2]) AND Data[3]) AND (NOT Data[4])) AND Data[23])) OR Data[19])) AND ((NOT ((((Data[1] AND Data[2]) AND Data[3]) AND (NOT Data[4])) AND Data[23])) OR Data[29])) AND ((NOT (((((NOT Data[1]) AND (NOT Data[2])) AND (NOT Data[3])) AND Data[4]) AND Data[23])) OR Data[30])) AND ((NOT ((((Data[1] AND (NOT Data[2])) AND (NOT Data[3])) AND Data[4]) AND Data[23])) OR Data[31])) AND ((NOT (((((NOT Data[1]) AND Data[2]) AND (NOT Data[3])) AND Data[4]) AND Data[23])) OR Data[32])) AND ((NOT ((((Data[1] AND Data[2]) AND (NOT Data[3])) AND Data[4]) AND Data[23])) OR Data[33])) AND ((NOT (((((NOT Data[1]) AND (NOT Data[2])) AND Data[3]) AND Data[4]) AND Data[23])) OR Data[34])) AND ((NOT ((((Data[1] AND (NOT Data[2])) AND Data[3]) AND Data[4]) AND Data[23])) OR Data[35])) AND ((NOT (((((NOT Data[1]) AND Data[2]) AND Data[3]) AND Data[4]) AND Data[23])) OR Data[36])) AND ((NOT ((((Data[1] AND Data[2]) AND Data[3]) AND Data[4]) AND Data[23])) OR Data[37]));
    OutReady := 1;
    CollectInput(RESET:=TRUE);
  END_IF;
END_PROGRAM

CONFIGURATION Config0
  RESOURCE Res0 ON PLC
    TASK task0(INTERVAL := T#20ms,PRIORITY := 0);
    PROGRAM instance0 WITH task0 : Boiler;
  END_RESOURCE
END_CONFIGURATION

(* ---- 5-MUX_warps-wield-plain.st ---- *)
(*
This code implements a shuffled multiplexer with 5 control bits.
The control bits are: Data[N1], Data[N22], Data[N24], Data[N20], Data[N21]
The input bits are: Data[N27], Data[N5], Data[N23], Data[N2], Data[N3], Data[N25], Data[N4], Data[N15], Data[N9], Data[N11], Data[N28], Data[N7], Data[N26], Data[N8], Data[N6], Data[N30], Data[N10], Data[N12], Data[N32], Data[N33], Data[N29], Data[N31], Data[N34], Data[N35], Data[N14], Data[N36], Data[N37], Data[N17], Data[N13], Data[N18], Data[N16], Data[N19]

The symbolic expression is:
((((((((((((((((((((((((((((((((!(((((!(IN1)) & (!(IN22))) & (!(IN24))) & (!(IN20))) & (!(IN21)))) | IN27) & ((!((((IN1 & (!(IN22))) & (!(IN24))) & (!(IN20))) & (!(IN21)))) | IN5)) & ((!(((((!(IN1)) & IN22) & (!(IN24))) & (!(IN20))) & (!(IN21)))) | IN23)) & ((!((((IN1 & IN22) & (!(IN24))) & (!(IN20))) & (!(IN21)))) | IN2)) & ((!(((((!(IN1)) & (!(IN22))) & IN24) & (!(IN20))) & (!(IN21)))) | IN3)) & ((!((((IN1 & (!(IN22))) & IN24) & (!(IN20))) & (!(IN21)))) | IN25)) & ((!(((((!(IN1)) & IN22) & IN24) & (!(IN20))) & (!(IN21)))) | IN4)) & ((!((((IN1 & IN22) & IN24) & (!(IN20))) & (!(IN21)))) | IN15)) & ((!(((((!(IN1)) & (!(IN22))) & (!(IN24))) & IN20) & (!(IN21)))) | IN9)) & ((!((((IN1 & (!(IN22))) & (!(IN24))) & IN20) & (!(IN21)))) | IN11)) & ((!(((((!(IN1)) & IN22) & (!(IN24))) & IN20) & (!(IN21)))) | IN28)) & ((!((((IN1 & IN22) & (!(IN24))) & IN20) & (!(IN21)))) | IN7)) & ((!(((((!(IN1)) & (!(IN22))) & IN24) & IN20) & (!(IN21)))) | IN26)) & ((!((((IN1 & (!(IN22))) & IN24) & IN20) & (!(IN21)))) | IN8)) & ((!(((((!(IN1)) & IN22) & IN24) & IN20) & (!(IN21)))) | IN6)) & ((!((((IN1 & IN22) & IN24) & IN20) & (!(IN21)))) | IN30)) & ((!(((((!(IN1)) & (!(IN22))) & (!(IN24))) & (!(IN20))) & IN21)) | IN10)) & ((!((((IN1 & (!(IN22))) & (!(IN24))) & (!(IN20))) & IN21)) | IN12)) & ((!(((((!(IN1)) & IN22) & (!(IN24))) & (!(IN20))) & IN21)) | IN32)) & ((!((((IN1 & IN22) & (!(IN24))) & (!(IN20))) & IN21)) | IN33)) & ((!(((((!(IN1)) & (!(IN22))) & IN24) & (!(IN20))) & IN21)) | IN29)) & ((!((((IN1 & (!(IN22))) & IN24) & (!(IN20))) & IN21)) | IN31)) & ((!(((((!(IN1)) & IN22) & IN24) & (!(IN20))) & IN21)) | IN34)) & ((!((((IN1 & IN22) & IN24) & (!(IN20))) & IN21)) | IN35)) & ((!(((((!(IN1)) & (!(IN22))) & (!(IN24))) & IN20) & IN21)) | IN14)) & ((!((((IN1 & (!(IN22))) & (!(IN24))) & IN20) & IN21)) | IN36)) & ((!(((((!(IN1)) & IN22) & (!(IN24))) & IN20) & IN21)) | IN37)) & ((!((((IN1 & IN22) & (!(IN24))) & IN20) & IN21)) | IN17)) & ((!(((((!(IN1)) & (!(IN22))) & IN24) & IN20) & IN21)) | IN13)) & ((!((((IN1 & (!(IN22))) & IN24) & IN20) & IN21)) | IN18)) & ((!(((((!(IN1)) & IN22) & IN24) & IN20) & IN21)) | IN16)) & ((!((((IN1 & IN22) & IN24) & IN20) & IN21)) | IN19)

*)

FUNCTION_BLOCK F_CollectInput
  VAR_IN_OUT
      Data : ARRAY[1..40] OF BOOL;
  END_VAR
  VAR_INPUT
      TICK  : BOOL := 0;
      IN1   : BOOL := 0;
      IN2   : BOOL := 0;
      IN3   : BOOL := 0;
      IN4   : BOOL := 0;
      IN5   : BOOL := 0;
      RESET : BOOL := FALSE;
  END_VAR
  VAR_OUTPUT
      Finished : BOOL;
  END_VAR
  VAR
      j    : USINT := 1;
      tock : BOOL  := 0;
  END_VAR
  IF NOT RESET AND tock = NOT TICK THEN
      Data[j]   := IN1;
      Data[j+1] := IN2;
      Data[j+2] := IN3;
      Data[j+3] := IN4;
      Data[j+4] := IN5;
      j := j + 5;
      tock := TICK;
  ELSE
      j := 1;
      tock := 0;
  END_IF;
  Finished := (j > 40);
END_FUNCTION_BLOCK

PROGRAM Boiler
  VAR
    Data  : ARRAY[1..40] OF BOOL;
    Ready : BOOL;
    CollectInput : F_CollectInput;
  END_VAR
  VAR
    TICK     AT %IX1.0 : BOOL;
    IN1      AT %IX0.3 : BOOL;
    IN2      AT %IX0.4 : BOOL;
    IN3      AT %IX0.5 : BOOL;
    IN4      AT %IX0.6 : BOOL;
    IN5      AT %IX0.7 : BOOL;
    OutReady AT %QX0.0 : BOOL := FALSE;
    FeedNext AT %QX0.1 : BOOL := FALSE;
    Out      AT %QX0.2 : BOOL;
  END_VAR
  CollectInput(TICK:=TICK, IN1:=IN1, IN2:=IN2, IN3:=IN3, IN4:=IN4, IN5:=IN5);
  Ready := CollectInput.Finished;
  FeedNext := 1;
  IF Ready THEN
    Out := (((((((((((((((((((((((((((((((((NOT (((((NOT Data[1]) AND (NOT Data[22])) AND (NOT Data[24])) AND (NOT Data[20])) AND (NOT Data[21]))) OR Data[27]) AND ((NOT ((((Data[1] AND (NOT Data[22])) AND (NOT Data[24])) AND (NOT Data[20])) AND (NOT Data[21]))) OR Data[5])) AND ((NOT (((((NOT Data[1]) AND Data[22]) AND (NOT Data[24])) AND (NOT Data[20])) AND (NOT Data[21]))) OR Data[23])) AND ((NOT ((((Data[1] AND Data[22]) AND (NOT Data[24])) AND (NOT Data[20])) AND (NOT Data[21]))) OR Data[2])) AND ((NOT (((((NOT Data[1]) AND (NOT Data[22])) AND Data[24]) AND (NOT Data[20])) AND (NOT Data[21]))) OR Data[3])) AND ((NOT ((((Data[1] AND (NOT Data[22])) AND Data[24]) AND (NOT Data[20])) AND (NOT Data[21]))) OR Data[25])) AND ((NOT (((((NOT Data[1]) AND Data[22]) AND Data[24]) AND (NOT Data[20])) AND (NOT Data[21]))) OR Data[4])) AND ((NOT ((((Data[1] AND Data[22]) AND Data[24]) AND (NOT Data[20])) AND (NOT Data[21]))) OR Data[15])) AND ((NOT (((((NOT Data[1]) AND (NOT Data[22])) AND (NOT Data[24])) AND Data[20]) AND (NOT Data[21]))) OR Data[9])) AND ((NOT ((((Data[1] AND (NOT Data[22])) AND (NOT Data[24])) AND Data[20]) AND (NOT Data[21]))) OR Data[11])) AND ((NOT (((((NOT Data[1]) AND Data[22]) AND (NOT Data[24])) AND Data[20]) AND (NOT Data[21]))) OR Data[28])) AND ((NOT ((((Data[1] AND Data[22]) AND (NOT Data[24])) AND Data[20]) AND (NOT Data[21]))) OR Data[7])) AND ((NOT (((((NOT Data[1]) AND (NOT Data[22])) AND Data[24]) AND Data[20]) AND (NOT Data[21]))) OR Data[26])) AND ((NOT ((((Data[1] AND (NOT Data[22])) AND Data[24]) AND Data[20]) AND (NOT Data[21]))) OR Data[8])) AND ((NOT (((((NOT Data[1]) AND Data[22]) AND Data[24]) AND Data[20]) AND (NOT Data[21]))) OR Data[6])) AND ((NOT ((((Data[1] AND Data[22]) AND Data[24]) AND Data[20]) AND (NOT Data[21]))) OR Data[30])) AND ((NOT (((((NOT Data[1]) AND (NOT Data[22])) AND (NOT Data[24])) AND (NOT Data[20])) AND Data[21])) OR Data[10])) AND ((NOT ((((Data[1] AND (NOT Data[22])) AND (NOT Data[24])) AND (NOT Data[20])) AND Data[21])) OR Data[12])) AND ((NOT (((((NOT Data[1]) AND Data[22]) AND (NOT Data[24])) AND (NOT Data[20])) AND Data[21])) OR Data[32])) AND ((NOT ((((Data[1] AND Data[22]) AND (NOT Data[24])) AND (NOT Data[20])) AND Data[21])) OR Data[33])) AND ((NOT (((((NOT Data[1]) AND (NOT Data[22])) AND Data[24]) AND (NOT Data[20])) AND Data[21])) OR Data[29])) AND ((NOT ((((Data[1] AND (NOT Data[22])) AND Data[24]) AND (NOT Data[20])) AND Data[21])) OR Data[31])) AND ((NOT (((((NOT Data[1]) AND Data[22]) AND Data[24]) AND (NOT Data[20])) AND Data[21])) OR Data[34])) AND ((NOT ((((Data[1] AND Data[22]) AND Data[24]) AND (NOT Data[20])) AND Data[21])) OR Data[35])) AND ((NOT (((((NOT Data[1]) AND (NOT Data[22])) AND (NOT Data[24])) AND Data[20]) AND Data[21])) OR Data[14])) AND ((NOT ((((Data[1] AND (NOT Data[22])) AND (NOT Data[24])) AND Data[20]) AND Data[21])) OR Data[36])) AND ((NOT (((((NOT Data[1]) AND Data[22]) AND (NOT Data[24])) AND Data[20]) AND Data[21])) OR Data[37])) AND ((NOT ((((Data[1] AND Data[22]) AND (NOT Data[24])) AND Data[20]) AND Data[21])) OR Data[17])) AND ((NOT (((((NOT Data[1]) AND (NOT Data[22])) AND Data[24]) AND Data[20]) AND Data[21])) OR Data[13])) AND ((NOT ((((Data[1] AND (NOT Data[22])) AND Data[24]) AND Data[20]) AND Data[21])) OR Data[18])) AND ((NOT (((((NOT Data[1]) AND Data[22]) AND Data[24]) AND Data[20]) AND Data[21])) OR Data[16])) AND ((NOT ((((Data[1] AND Data[22]) AND Data[24]) AND Data[20]) AND Data[21])) OR Data[19]));
    OutReady := 1;
    CollectInput(RESET:=TRUE);
  END_IF;
END_PROGRAM

CONFIGURATION Config0
  RESOURCE Res0 ON PLC
    TASK task0(INTERVAL := T#20ms,PRIORITY := 0);
    PROGRAM instance0 WITH task0 : Boiler;
  END_RESOURCE
END_CONFIGURATION

(* ---- 5-MUX_wasps-image-petri.st ---- *)
(*
This code implements a shuffled multiplexer with 5 control bits.
The control bits are: Data[N1], Data[N2], Data[N23], Data[N3], Data[N22]
The input bits are: Data[N25], Data[N4], Data[N24], Data[N5], Data[N21], Data[N6], Data[N11], Data[N20], Data[N7], Data[N8], Data[N9], Data[N28], Data[N10], Data[N13], Data[N14], Data[N15], Data[N12], Data[N26], Data[N29], Data[N30], Data[N16], Data[N19], Data[N17], Data[N31], Data[N32], Data[N33], Data[N27], Data[N18], Data[N34], Data[N37], Data[N35], Data[N36]

The symbolic expression is:
((((((((((((((((((((((((((((((((!(((((!(IN1)) & (!(IN2))) & (!(IN23))) & (!(IN3))) & (!(IN22)))) | IN25) & ((!((((IN1 & (!(IN2))) & (!(IN23))) & (!(IN3))) & (!(IN22)))) | IN4)) & ((!(((((!(IN1)) & IN2) & (!(IN23))) & (!(IN3))) & (!(IN22)))) | IN24)) & ((!((((IN1 & IN2) & (!(IN23))) & (!(IN3))) & (!(IN22)))) | IN5)) & ((!(((((!(IN1)) & (!(IN2))) & IN23) & (!(IN3))) & (!(IN22)))) | IN21)) & ((!((((IN1 & (!(IN2))) & IN23) & (!(IN3))) & (!(IN22)))) | IN6)) & ((!(((((!(IN1)) & IN2) & IN23) & (!(IN3))) & (!(IN22)))) | IN11)) & ((!((((IN1 & IN2) & IN23) & (!(IN3))) & (!(IN22)))) | IN20)) & ((!(((((!(IN1)) & (!(IN2))) & (!(IN23))) & IN3) & (!(IN22)))) | IN7)) & ((!((((IN1 & (!(IN2))) & (!(IN23))) & IN3) & (!(IN22)))) | IN8)) & ((!(((((!(IN1)) & IN2) & (!(IN23))) & IN3) & (!(IN22)))) | IN9)) & ((!((((IN1 & IN2) & (!(IN23))) & IN3) & (!(IN22)))) | IN28)) & ((!(((((!(IN1)) & (!(IN2))) & IN23) & IN3) & (!(IN22)))) | IN10)) & ((!((((IN1 & (!(IN2))) & IN23) & IN3) & (!(IN22)))) | IN13)) & ((!(((((!(IN1)) & IN2) & IN23) & IN3) & (!(IN22)))) | IN14)) & ((!((((IN1 & IN2) & IN23) & IN3) & (!(IN22)))) | IN15)) & ((!(((((!(IN1)) & (!(IN2))) & (!(IN23))) & (!(IN3))) & IN22)) | IN12)) & ((!((((IN1 & (!(IN2))) & (!(IN23))) & (!(IN3))) & IN22)) | IN26)) & ((!(((((!(IN1)) & IN2) & (!(IN23))) & (!(IN3))) & IN22)) | IN29)) & ((!((((IN1 & IN2) & (!(IN23))) & (!(IN3))) & IN22)) | IN30)) & ((!(((((!(IN1)) & (!(IN2))) & IN23) & (!(IN3))) & IN22)) | IN16)) & ((!((((IN1 & (!(IN2))) & IN23) & (!(IN3))) & IN22)) | IN19)) & ((!(((((!(IN1)) & IN2) & IN23) & (!(IN3))) & IN22)) | IN17)) & ((!((((IN1 & IN2) & IN23) & (!(IN3))) & IN22)) | IN31)) & ((!(((((!(IN1)) & (!(IN2))) & (!(IN23))) & IN3) & IN22)) | IN32)) & ((!((((IN1 & (!(IN2))) & (!(IN23))) & IN3) & IN22)) | IN33)) & ((!(((((!(IN1)) & IN2) & (!(IN23))) & IN3) & IN22)) | IN27)) & ((!((((IN1 & IN2) & (!(IN23))) & IN3) & IN22)) | IN18)) & ((!(((((!(IN1)) & (!(IN2))) & IN23) & IN3) & IN22)) | IN34)) & ((!((((IN1 & (!(IN2))) & IN23) & IN3) & IN22)) | IN37)) & ((!(((((!(IN1)) & IN2) & IN23) & IN3) & IN22)) | IN35)) & ((!((((IN1 & IN2) & IN23) & IN3) & IN22)) | IN36)

*)

FUNCTION_BLOCK F_CollectInput
  VAR_IN_OUT
      Data : ARRAY[1..40] OF BOOL;
  END_VAR
  VAR_INPUT
      TICK  : BOOL := 0;
      IN1   : BOOL := 0;
      IN2   : BOOL := 0;
      IN3   : BOOL := 0;
      IN4   : BOOL := 0;
      IN5   : BOOL := 0;
      RESET : BOOL := FALSE;
  END_VAR
  VAR_OUTPUT
      Finished : BOOL;
  END_VAR
  VAR
      j    : USINT := 1;
      tock : BOOL  := 0;
  END_VAR
  IF NOT RESET AND tock = NOT TICK THEN
      Data[j]   := IN1;
      Data[j+1] := IN2;
      Data[j+2] := IN3;
      Data[j+3] := IN4;
      Data[j+4] := IN5;
      j := j + 5;
      tock := TICK;
  ELSE
      j := 1;
      tock := 0;
  END_IF;
  Finished := (j > 40);
END_FUNCTION_BLOCK

PROGRAM Boiler
  VAR
    Data  : ARRAY[1..40] OF BOOL;
    Ready : BOOL;
    CollectInput : F_CollectInput;
  END_VAR
  VAR
    TICK     AT %IX1.0 : BOOL;
    IN1      AT %IX0.3 : BOOL;
    IN2      AT %IX0.4 : BOOL;
    IN3      AT %IX0.5 : BOOL;
    IN4      AT %IX0.6 : BOOL;
    IN5      AT %IX0.7 : BOOL;
    OutReady AT %QX0.0 : BOOL := FALSE;
    FeedNext AT %QX0.1 : BOOL := FALSE;
    Out      AT %QX0.2 : BOOL;
  END_VAR
  CollectInput(TICK:=TICK, IN1:=IN1, IN2:=IN2, IN3:=IN3, IN4:=IN4, IN5:=IN5);
  Ready := CollectInput.Finished;
  FeedNext := 1;
  IF Ready THEN
    Out := (((((((((((((((((((((((((((((((((NOT (((((NOT Data[1]) AND (NOT Data[2])) AND (NOT Data[23])) AND (NOT Data[3])) AND (NOT Data[22]))) OR Data[25]) AND ((NOT ((((Data[1] AND (NOT Data[2])) AND (NOT Data[23])) AND (NOT Data[3])) AND (NOT Data[22]))) OR Data[4])) AND ((NOT (((((NOT Data[1]) AND Data[2]) AND (NOT Data[23])) AND (NOT Data[3])) AND (NOT Data[22]))) OR Data[24])) AND ((NOT ((((Data[1] AND Data[2]) AND (NOT Data[23])) AND (NOT Data[3])) AND (NOT Data[22]))) OR Data[5])) AND ((NOT (((((NOT Data[1]) AND (NOT Data[2])) AND Data[23]) AND (NOT Data[3])) AND (NOT Data[22]))) OR Data[21])) AND ((NOT ((((Data[1] AND (NOT Data[2])) AND Data[23]) AND (NOT Data[3])) AND (NOT Data[22]))) OR Data[6])) AND ((NOT (((((NOT Data[1]) AND Data[2]) AND Data[23]) AND (NOT Data[3])) AND (NOT Data[22]))) OR Data[11])) AND ((NOT ((((Data[1] AND Data[2]) AND Data[23]) AND (NOT Data[3])) AND (NOT Data[22]))) OR Data[20])) AND ((NOT (((((NOT Data[1]) AND (NOT Data[2])) AND (NOT Data[23])) AND Data[3]) AND (NOT Data[22]))) OR Data[7])) AND ((NOT ((((Data[1] AND (NOT Data[2])) AND (NOT Data[23])) AND Data[3]) AND (NOT Data[22]))) OR Data[8])) AND ((NOT (((((NOT Data[1]) AND Data[2]) AND (NOT Data[23])) AND Data[3]) AND (NOT Data[22]))) OR Data[9])) AND ((NOT ((((Data[1] AND Data[2]) AND (NOT Data[23])) AND Data[3]) AND (NOT Data[22]))) OR Data[28])) AND ((NOT (((((NOT Data[1]) AND (NOT Data[2])) AND Data[23]) AND Data[3]) AND (NOT Data[22]))) OR Data[10])) AND ((NOT ((((Data[1] AND (NOT Data[2])) AND Data[23]) AND Data[3]) AND (NOT Data[22]))) OR Data[13])) AND ((NOT (((((NOT Data[1]) AND Data[2]) AND Data[23]) AND Data[3]) AND (NOT Data[22]))) OR Data[14])) AND ((NOT ((((Data[1] AND Data[2]) AND Data[23]) AND Data[3]) AND (NOT Data[22]))) OR Data[15])) AND ((NOT (((((NOT Data[1]) AND (NOT Data[2])) AND (NOT Data[23])) AND (NOT Data[3])) AND Data[22])) OR Data[12])) AND ((NOT ((((Data[1] AND (NOT Data[2])) AND (NOT Data[23])) AND (NOT Data[3])) AND Data[22])) OR Data[26])) AND ((NOT (((((NOT Data[1]) AND Data[2]) AND (NOT Data[23])) AND (NOT Data[3])) AND Data[22])) OR Data[29])) AND ((NOT ((((Data[1] AND Data[2]) AND (NOT Data[23])) AND (NOT Data[3])) AND Data[22])) OR Data[30])) AND ((NOT (((((NOT Data[1]) AND (NOT Data[2])) AND Data[23]) AND (NOT Data[3])) AND Data[22])) OR Data[16])) AND ((NOT ((((Data[1] AND (NOT Data[2])) AND Data[23]) AND (NOT Data[3])) AND Data[22])) OR Data[19])) AND ((NOT (((((NOT Data[1]) AND Data[2]) AND Data[23]) AND (NOT Data[3])) AND Data[22])) OR Data[17])) AND ((NOT ((((Data[1] AND Data[2]) AND Data[23]) AND (NOT Data[3])) AND Data[22])) OR Data[31])) AND ((NOT (((((NOT Data[1]) AND (NOT Data[2])) AND (NOT Data[23])) AND Data[3]) AND Data[22])) OR Data[32])) AND ((NOT ((((Data[1] AND (NOT Data[2])) AND (NOT Data[23])) AND Data[3]) AND Data[22])) OR Data[33])) AND ((NOT (((((NOT Data[1]) AND Data[2]) AND (NOT Data[23])) AND Data[3]) AND Data[22])) OR Data[27])) AND ((NOT ((((Data[1] AND Data[2]) AND (NOT Data[23])) AND Data[3]) AND Data[22])) OR Data[18])) AND ((NOT (((((NOT Data[1]) AND (NOT Data[2])) AND Data[23]) AND Data[3]) AND Data[22])) OR Data[34])) AND ((NOT ((((Data[1] AND (NOT Data[2])) AND Data[23]) AND Data[3]) AND Data[22])) OR Data[37])) AND ((NOT (((((NOT Data[1]) AND Data[2]) AND Data[23]) AND Data[3]) AND Data[22])) OR Data[35])) AND ((NOT ((((Data[1] AND Data[2]) AND Data[23]) AND Data[3]) AND Data[22])) OR Data[36]));
    OutReady := 1;
    CollectInput(RESET:=TRUE);
  END_IF;
END_PROGRAM

CONFIGURATION Config0
  RESOURCE Res0 ON PLC
    TASK task0(INTERVAL := T#20ms,PRIORITY := 0);
    PROGRAM instance0 WITH task0 : Boiler;
  END_RESOURCE
END_CONFIGURATION

(* ---- 5-MUX_waved-cocoa-undid.st ---- *)
(*
This code implements a shuffled multiplexer with 5 control bits.
The control bits are: Data[N27], Data[N1], Data[N2], Data[N3], Data[N23]
The input bits are: Data[N4], Data[N22], Data[N20], Data[N10], Data[N5], Data[N12], Data[N24], Data[N8], Data[N6], Data[N26], Data[N7], Data[N11], Data[N13], Data[N32], Data[N9], Data[N14], Data[N18], Data[N21], Data[N33], Data[N15], Data[N25], Data[N28], Data[N16], Data[N17], Data[N30], Data[N19], Data[N29], Data[N35], Data[N31], Data[N34], Data[N36], Data[N37]

The symbolic expression is:
((((((((((((((((((((((((((((((((!(((((!(IN27)) & (!(IN1))) & (!(IN2))) & (!(IN3))) & (!(IN23)))) | IN4) & ((!((((IN27 & (!(IN1))) & (!(IN2))) & (!(IN3))) & (!(IN23)))) | IN22)) & ((!(((((!(IN27)) & IN1) & (!(IN2))) & (!(IN3))) & (!(IN23)))) | IN20)) & ((!((((IN27 & IN1) & (!(IN2))) & (!(IN3))) & (!(IN23)))) | IN10)) & ((!(((((!(IN27)) & (!(IN1))) & IN2) & (!(IN3))) & (!(IN23)))) | IN5)) & ((!((((IN27 & (!(IN1))) & IN2) & (!(IN3))) & (!(IN23)))) | IN12)) & ((!(((((!(IN27)) & IN1) & IN2) & (!(IN3))) & (!(IN23)))) | IN24)) & ((!((((IN27 & IN1) & IN2) & (!(IN3))) & (!(IN23)))) | IN8)) & ((!(((((!(IN27)) & (!(IN1))) & (!(IN2))) & IN3) & (!(IN23)))) | IN6)) & ((!((((IN27 & (!(IN1))) & (!(IN2))) & IN3) & (!(IN23)))) | IN26)) & ((!(((((!(IN27)) & IN1) & (!(IN2))) & IN3) & (!(IN23)))) | IN7)) & ((!((((IN27 & IN1) & (!(IN2))) & IN3) & (!(IN23)))) | IN11)) & ((!(((((!(IN27)) & (!(IN1))) & IN2) & IN3) & (!(IN23)))) | IN13)) & ((!((((IN27 & (!(IN1))) & IN2) & IN3) & (!(IN23)))) | IN32)) & ((!(((((!(IN27)) & IN1) & IN2) & IN3) & (!(IN23)))) | IN9)) & ((!((((IN27 & IN1) & IN2) & IN3) & (!(IN23)))) | IN14)) & ((!(((((!(IN27)) & (!(IN1))) & (!(IN2))) & (!(IN3))) & IN23)) | IN18)) & ((!((((IN27 & (!(IN1))) & (!(IN2))) & (!(IN3))) & IN23)) | IN21)) & ((!(((((!(IN27)) & IN1) & (!(IN2))) & (!(IN3))) & IN23)) | IN33)) & ((!((((IN27 & IN1) & (!(IN2))) & (!(IN3))) & IN23)) | IN15)) & ((!(((((!(IN27)) & (!(IN1))) & IN2) & (!(IN3))) & IN23)) | IN25)) & ((!((((IN27 & (!(IN1))) & IN2) & (!(IN3))) & IN23)) | IN28)) & ((!(((((!(IN27)) & IN1) & IN2) & (!(IN3))) & IN23)) | IN16)) & ((!((((IN27 & IN1) & IN2) & (!(IN3))) & IN23)) | IN17)) & ((!(((((!(IN27)) & (!(IN1))) & (!(IN2))) & IN3) & IN23)) | IN30)) & ((!((((IN27 & (!(IN1))) & (!(IN2))) & IN3) & IN23)) | IN19)) & ((!(((((!(IN27)) & IN1) & (!(IN2))) & IN3) & IN23)) | IN29)) & ((!((((IN27 & IN1) & (!(IN2))) & IN3) & IN23)) | IN35)) & ((!(((((!(IN27)) & (!(IN1))) & IN2) & IN3) & IN23)) | IN31)) & ((!((((IN27 & (!(IN1))) & IN2) & IN3) & IN23)) | IN34)) & ((!(((((!(IN27)) & IN1) & IN2) & IN3) & IN23)) | IN36)) & ((!((((IN27 & IN1) & IN2) & IN3) & IN23)) | IN37)

*)

FUNCTION_BLOCK F_CollectInput
  VAR_IN_OUT
      Data : ARRAY[1..40] OF BOOL;
  END_VAR
  VAR_INPUT
      TICK  : BOOL := 0;
      IN1   : BOOL := 0;
      IN2   : BOOL := 0;
      IN3   : BOOL := 0;
      IN4   : BOOL := 0;
      IN5   : BOOL := 0;
      RESET : BOOL := FALSE;
  END_VAR
  VAR_OUTPUT
      Finished : BOOL;
  END_VAR
  VAR
      j    : USINT := 1;
      tock : BOOL  := 0;
  END_VAR
  IF NOT RESET AND tock = NOT TICK THEN
      Data[j]   := IN1;
      Data[j+1] := IN2;
      Data[j+2] := IN3;
      Data[j+3] := IN4;
      Data[j+4] := IN5;
      j := j + 5;
      tock := TICK;
  ELSE
      j := 1;
      tock := 0;
  END_IF;
  Finished := (j > 40);
END_FUNCTION_BLOCK

PROGRAM Boiler
  VAR
    Data  : ARRAY[1..40] OF BOOL;
    Ready : BOOL;
    CollectInput : F_CollectInput;
  END_VAR
  VAR
    TICK     AT %IX1.0 : BOOL;
    IN1      AT %IX0.3 : BOOL;
    IN2      AT %IX0.4 : BOOL;
    IN3      AT %IX0.5 : BOOL;
    IN4      AT %IX0.6 : BOOL;
    IN5      AT %IX0.7 : BOOL;
    OutReady AT %QX0.0 : BOOL := FALSE;
    FeedNext AT %QX0.1 : BOOL := FALSE;
    Out      AT %QX0.2 : BOOL;
  END_VAR
  CollectInput(TICK:=TICK, IN1:=IN1, IN2:=IN2, IN3:=IN3, IN4:=IN4, IN5:=IN5);
  Ready := CollectInput.Finished;
  FeedNext := 1;
  IF Ready THEN
    Out := (((((((((((((((((((((((((((((((((NOT (((((NOT Data[27]) AND (NOT Data[1])) AND (NOT Data[2])) AND (NOT Data[3])) AND (NOT Data[23]))) OR Data[4]) AND ((NOT ((((Data[27] AND (NOT Data[1])) AND (NOT Data[2])) AND (NOT Data[3])) AND (NOT Data[23]))) OR Data[22])) AND ((NOT (((((NOT Data[27]) AND Data[1]) AND (NOT Data[2])) AND (NOT Data[3])) AND (NOT Data[23]))) OR Data[20])) AND ((NOT ((((Data[27] AND Data[1]) AND (NOT Data[2])) AND (NOT Data[3])) AND (NOT Data[23]))) OR Data[10])) AND ((NOT (((((NOT Data[27]) AND (NOT Data[1])) AND Data[2]) AND (NOT Data[3])) AND (NOT Data[23]))) OR Data[5])) AND ((NOT ((((Data[27] AND (NOT Data[1])) AND Data[2]) AND (NOT Data[3])) AND (NOT Data[23]))) OR Data[12])) AND ((NOT (((((NOT Data[27]) AND Data[1]) AND Data[2]) AND (NOT Data[3])) AND (NOT Data[23]))) OR Data[24])) AND ((NOT ((((Data[27] AND Data[1]) AND Data[2]) AND (NOT Data[3])) AND (NOT Data[23]))) OR Data[8])) AND ((NOT (((((NOT Data[27]) AND (NOT Data[1])) AND (NOT Data[2])) AND Data[3]) AND (NOT Data[23]))) OR Data[6])) AND ((NOT ((((Data[27] AND (NOT Data[1])) AND (NOT Data[2])) AND Data[3]) AND (NOT Data[23]))) OR Data[26])) AND ((NOT (((((NOT Data[27]) AND Data[1]) AND (NOT Data[2])) AND Data[3]) AND (NOT Data[23]))) OR Data[7])) AND ((NOT ((((Data[27] AND Data[1]) AND (NOT Data[2])) AND Data[3]) AND (NOT Data[23]))) OR Data[11])) AND ((NOT (((((NOT Data[27]) AND (NOT Data[1])) AND Data[2]) AND Data[3]) AND (NOT Data[23]))) OR Data[13])) AND ((NOT ((((Data[27] AND (NOT Data[1])) AND Data[2]) AND Data[3]) AND (NOT Data[23]))) OR Data[32])) AND ((NOT (((((NOT Data[27]) AND Data[1]) AND Data[2]) AND Data[3]) AND (NOT Data[23]))) OR Data[9])) AND ((NOT ((((Data[27] AND Data[1]) AND Data[2]) AND Data[3]) AND (NOT Data[23]))) OR Data[14])) AND ((NOT (((((NOT Data[27]) AND (NOT Data[1])) AND (NOT Data[2])) AND (NOT Data[3])) AND Data[23])) OR Data[18])) AND ((NOT ((((Data[27] AND (NOT Data[1])) AND (NOT Data[2])) AND (NOT Data[3])) AND Data[23])) OR Data[21])) AND ((NOT (((((NOT Data[27]) AND Data[1]) AND (NOT Data[2])) AND (NOT Data[3])) AND Data[23])) OR Data[33])) AND ((NOT ((((Data[27] AND Data[1]) AND (NOT Data[2])) AND (NOT Data[3])) AND Data[23])) OR Data[15])) AND ((NOT (((((NOT Data[27]) AND (NOT Data[1])) AND Data[2]) AND (NOT Data[3])) AND Data[23])) OR Data[25])) AND ((NOT ((((Data[27] AND (NOT Data[1])) AND Data[2]) AND (NOT Data[3])) AND Data[23])) OR Data[28])) AND ((NOT (((((NOT Data[27]) AND Data[1]) AND Data[2]) AND (NOT Data[3])) AND Data[23])) OR Data[16])) AND ((NOT ((((Data[27] AND Data[1]) AND Data[2]) AND (NOT Data[3])) AND Data[23])) OR Data[17])) AND ((NOT (((((NOT Data[27]) AND (NOT Data[1])) AND (NOT Data[2])) AND Data[3]) AND Data[23])) OR Data[30])) AND ((NOT ((((Data[27] AND (NOT Data[1])) AND (NOT Data[2])) AND Data[3]) AND Data[23])) OR Data[19])) AND ((NOT (((((NOT Data[27]) AND Data[1]) AND (NOT Data[2])) AND Data[3]) AND Data[23])) OR Data[29])) AND ((NOT ((((Data[27] AND Data[1]) AND (NOT Data[2])) AND Data[3]) AND Data[23])) OR Data[35])) AND ((NOT (((((NOT Data[27]) AND (NOT Data[1])) AND Data[2]) AND Data[3]) AND Data[23])) OR Data[31])) AND ((NOT ((((Data[27] AND (NOT Data[1])) AND Data[2]) AND Data[3]) AND Data[23])) OR Data[34])) AND ((NOT (((((NOT Data[27]) AND Data[1]) AND Data[2]) AND Data[3]) AND Data[23])) OR Data[36])) AND ((NOT ((((Data[27] AND Data[1]) AND Data[2]) AND Data[3]) AND Data[23])) OR Data[37]));
    OutReady := 1;
    CollectInput(RESET:=TRUE);
  END_IF;
END_PROGRAM

CONFIGURATION Config0
  RESOURCE Res0 ON PLC
    TASK task0(INTERVAL := T#20ms,PRIORITY := 0);
    PROGRAM instance0 WITH task0 : Boiler;
  END_RESOURCE
END_CONFIGURATION

(* ---- 5-MUX_wench-khans-fasts.st ---- *)
(*
This code implements a shuffled multiplexer with 5 control bits.
The control bits are: Data[N1], Data[N2], Data[N3], Data[N22], Data[N23]
The input bits are: Data[N4], Data[N21], Data[N20], Data[N26], Data[N28], Data[N29], Data[N6], Data[N5], Data[N7], Data[N8], Data[N9], Data[N27], Data[N12], Data[N10], Data[N31], Data[N13], Data[N11], Data[N24], Data[N30], Data[N14], Data[N16], Data[N35], Data[N25], Data[N17], Data[N19], Data[N32], Data[N15], Data[N33], Data[N34], Data[N36], Data[N18], Data[N37]

The symbolic expression is:
((((((((((((((((((((((((((((((((!(((((!(IN1)) & (!(IN2))) & (!(IN3))) & (!(IN22))) & (!(IN23)))) | IN4) & ((!((((IN1 & (!(IN2))) & (!(IN3))) & (!(IN22))) & (!(IN23)))) | IN21)) & ((!(((((!(IN1)) & IN2) & (!(IN3))) & (!(IN22))) & (!(IN23)))) | IN20)) & ((!((((IN1 & IN2) & (!(IN3))) & (!(IN22))) & (!(IN23)))) | IN26)) & ((!(((((!(IN1)) & (!(IN2))) & IN3) & (!(IN22))) & (!(IN23)))) | IN28)) & ((!((((IN1 & (!(IN2))) & IN3) & (!(IN22))) & (!(IN23)))) | IN29)) & ((!(((((!(IN1)) & IN2) & IN3) & (!(IN22))) & (!(IN23)))) | IN6)) & ((!((((IN1 & IN2) & IN3) & (!(IN22))) & (!(IN23)))) | IN5)) & ((!(((((!(IN1)) & (!(IN2))) & (!(IN3))) & IN22) & (!(IN23)))) | IN7)) & ((!((((IN1 & (!(IN2))) & (!(IN3))) & IN22) & (!(IN23)))) | IN8)) & ((!(((((!(IN1)) & IN2) & (!(IN3))) & IN22) & (!(IN23)))) | IN9)) & ((!((((IN1 & IN2) & (!(IN3))) & IN22) & (!(IN23)))) | IN27)) & ((!(((((!(IN1)) & (!(IN2))) & IN3) & IN22) & (!(IN23)))) | IN12)) & ((!((((IN1 & (!(IN2))) & IN3) & IN22) & (!(IN23)))) | IN10)) & ((!(((((!(IN1)) & IN2) & IN3) & IN22) & (!(IN23)))) | IN31)) & ((!((((IN1 & IN2) & IN3) & IN22) & (!(IN23)))) | IN13)) & ((!(((((!(IN1)) & (!(IN2))) & (!(IN3))) & (!(IN22))) & IN23)) | IN11)) & ((!((((IN1 & (!(IN2))) & (!(IN3))) & (!(IN22))) & IN23)) | IN24)) & ((!(((((!(IN1)) & IN2) & (!(IN3))) & (!(IN22))) & IN23)) | IN30)) & ((!((((IN1 & IN2) & (!(IN3))) & (!(IN22))) & IN23)) | IN14)) & ((!(((((!(IN1)) & (!(IN2))) & IN3) & (!(IN22))) & IN23)) | IN16)) & ((!((((IN1 & (!(IN2))) & IN3) & (!(IN22))) & IN23)) | IN35)) & ((!(((((!(IN1)) & IN2) & IN3) & (!(IN22))) & IN23)) | IN25)) & ((!((((IN1 & IN2) & IN3) & (!(IN22))) & IN23)) | IN17)) & ((!(((((!(IN1)) & (!(IN2))) & (!(IN3))) & IN22) & IN23)) | IN19)) & ((!((((IN1 & (!(IN2))) & (!(IN3))) & IN22) & IN23)) | IN32)) & ((!(((((!(IN1)) & IN2) & (!(IN3))) & IN22) & IN23)) | IN15)) & ((!((((IN1 & IN2) & (!(IN3))) & IN22) & IN23)) | IN33)) & ((!(((((!(IN1)) & (!(IN2))) & IN3) & IN22) & IN23)) | IN34)) & ((!((((IN1 & (!(IN2))) & IN3) & IN22) & IN23)) | IN36)) & ((!(((((!(IN1)) & IN2) & IN3) & IN22) & IN23)) | IN18)) & ((!((((IN1 & IN2) & IN3) & IN22) & IN23)) | IN37)

*)

FUNCTION_BLOCK F_CollectInput
  VAR_IN_OUT
      Data : ARRAY[1..40] OF BOOL;
  END_VAR
  VAR_INPUT
      TICK  : BOOL := 0;
      IN1   : BOOL := 0;
      IN2   : BOOL := 0;
      IN3   : BOOL := 0;
      IN4   : BOOL := 0;
      IN5   : BOOL := 0;
      RESET : BOOL := FALSE;
  END_VAR
  VAR_OUTPUT
      Finished : BOOL;
  END_VAR
  VAR
      j    : USINT := 1;
      tock : BOOL  := 0;
  END_VAR
  IF NOT RESET AND tock = NOT TICK THEN
      Data[j]   := IN1;
      Data[j+1] := IN2;
      Data[j+2] := IN3;
      Data[j+3] := IN4;
      Data[j+4] := IN5;
      j := j + 5;
      tock := TICK;
  ELSE
      j := 1;
      tock := 0;
  END_IF;
  Finished := (j > 40);
END_FUNCTION_BLOCK

PROGRAM Boiler
  VAR
    Data  : ARRAY[1..40] OF BOOL;
    Ready : BOOL;
    CollectInput : F_CollectInput;
  END_VAR
  VAR
    TICK     AT %IX1.0 : BOOL;
    IN1      AT %IX0.3 : BOOL;
    IN2      AT %IX0.4 : BOOL;
    IN3      AT %IX0.5 : BOOL;
    IN4      AT %IX0.6 : BOOL;
    IN5      AT %IX0.7 : BOOL;
    OutReady AT %QX0.0 : BOOL := FALSE;
    FeedNext AT %QX0.1 : BOOL := FALSE;
    Out      AT %QX0.2 : BOOL;
  END_VAR
  CollectInput(TICK:=TICK, IN1:=IN1, IN2:=IN2, IN3:=IN3, IN4:=IN4, IN5:=IN5);
  Ready := CollectInput.Finished;
  FeedNext := 1;
  IF Ready THEN
    Out := (((((((((((((((((((((((((((((((((NOT (((((NOT Data[1]) AND (NOT Data[2])) AND (NOT Data[3])) AND (NOT Data[22])) AND (NOT Data[23]))) OR Data[4]) AND ((NOT ((((Data[1] AND (NOT Data[2])) AND (NOT Data[3])) AND (NOT Data[22])) AND (NOT Data[23]))) OR Data[21])) AND ((NOT (((((NOT Data[1]) AND Data[2]) AND (NOT Data[3])) AND (NOT Data[22])) AND (NOT Data[23]))) OR Data[20])) AND ((NOT ((((Data[1] AND Data[2]) AND (NOT Data[3])) AND (NOT Data[22])) AND (NOT Data[23]))) OR Data[26])) AND ((NOT (((((NOT Data[1]) AND (NOT Data[2])) AND Data[3]) AND (NOT Data[22])) AND (NOT Data[23]))) OR Data[28])) AND ((NOT ((((Data[1] AND (NOT Data[2])) AND Data[3]) AND (NOT Data[22])) AND (NOT Data[23]))) OR Data[29])) AND ((NOT (((((NOT Data[1]) AND Data[2]) AND Data[3]) AND (NOT Data[22])) AND (NOT Data[23]))) OR Data[6])) AND ((NOT ((((Data[1] AND Data[2]) AND Data[3]) AND (NOT Data[22])) AND (NOT Data[23]))) OR Data[5])) AND ((NOT (((((NOT Data[1]) AND (NOT Data[2])) AND (NOT Data[3])) AND Data[22]) AND (NOT Data[23]))) OR Data[7])) AND ((NOT ((((Data[1] AND (NOT Data[2])) AND (NOT Data[3])) AND Data[22]) AND (NOT Data[23]))) OR Data[8])) AND ((NOT (((((NOT Data[1]) AND Data[2]) AND (NOT Data[3])) AND Data[22]) AND (NOT Data[23]))) OR Data[9])) AND ((NOT ((((Data[1] AND Data[2]) AND (NOT Data[3])) AND Data[22]) AND (NOT Data[23]))) OR Data[27])) AND ((NOT (((((NOT Data[1]) AND (NOT Data[2])) AND Data[3]) AND Data[22]) AND (NOT Data[23]))) OR Data[12])) AND ((NOT ((((Data[1] AND (NOT Data[2])) AND Data[3]) AND Data[22]) AND (NOT Data[23]))) OR Data[10])) AND ((NOT (((((NOT Data[1]) AND Data[2]) AND Data[3]) AND Data[22]) AND (NOT Data[23]))) OR Data[31])) AND ((NOT ((((Data[1] AND Data[2]) AND Data[3]) AND Data[22]) AND (NOT Data[23]))) OR Data[13])) AND ((NOT (((((NOT Data[1]) AND (NOT Data[2])) AND (NOT Data[3])) AND (NOT Data[22])) AND Data[23])) OR Data[11])) AND ((NOT ((((Data[1] AND (NOT Data[2])) AND (NOT Data[3])) AND (NOT Data[22])) AND Data[23])) OR Data[24])) AND ((NOT (((((NOT Data[1]) AND Data[2]) AND (NOT Data[3])) AND (NOT Data[22])) AND Data[23])) OR Data[30])) AND ((NOT ((((Data[1] AND Data[2]) AND (NOT Data[3])) AND (NOT Data[22])) AND Data[23])) OR Data[14])) AND ((NOT (((((NOT Data[1]) AND (NOT Data[2])) AND Data[3]) AND (NOT Data[22])) AND Data[23])) OR Data[16])) AND ((NOT ((((Data[1] AND (NOT Data[2])) AND Data[3]) AND (NOT Data[22])) AND Data[23])) OR Data[35])) AND ((NOT (((((NOT Data[1]) AND Data[2]) AND Data[3]) AND (NOT Data[22])) AND Data[23])) OR Data[25])) AND ((NOT ((((Data[1] AND Data[2]) AND Data[3]) AND (NOT Data[22])) AND Data[23])) OR Data[17])) AND ((NOT (((((NOT Data[1]) AND (NOT Data[2])) AND (NOT Data[3])) AND Data[22]) AND Data[23])) OR Data[19])) AND ((NOT ((((Data[1] AND (NOT Data[2])) AND (NOT Data[3])) AND Data[22]) AND Data[23])) OR Data[32])) AND ((NOT (((((NOT Data[1]) AND Data[2]) AND (NOT Data[3])) AND Data[22]) AND Data[23])) OR Data[15])) AND ((NOT ((((Data[1] AND Data[2]) AND (NOT Data[3])) AND Data[22]) AND Data[23])) OR Data[33])) AND ((NOT (((((NOT Data[1]) AND (NOT Data[2])) AND Data[3]) AND Data[22]) AND Data[23])) OR Data[34])) AND ((NOT ((((Data[1] AND (NOT Data[2])) AND Data[3]) AND Data[22]) AND Data[23])) OR Data[36])) AND ((NOT (((((NOT Data[1]) AND Data[2]) AND Data[3]) AND Data[22]) AND Data[23])) OR Data[18])) AND ((NOT ((((Data[1] AND Data[2]) AND Data[3]) AND Data[22]) AND Data[23])) OR Data[37]));
    OutReady := 1;
    CollectInput(RESET:=TRUE);
  END_IF;
END_PROGRAM

CONFIGURATION Config0
  RESOURCE Res0 ON PLC
    TASK task0(INTERVAL := T#20ms,PRIORITY := 0);
    PROGRAM instance0 WITH task0 : Boiler;
  END_RESOURCE
END_CONFIGURATION

(* ---- 5-MUX_world-maced-wings.st ---- *)
(*
This code implements a shuffled multiplexer with 5 control bits.
The control bits are: Data[N4], Data[N2], Data[N22], Data[N3], Data[N21]
The input bits are: Data[N1], Data[N5], Data[N20], Data[N7], Data[N6], Data[N8], Data[N23], Data[N10], Data[N26], Data[N28], Data[N25], Data[N27], Data[N12], Data[N30], Data[N24], Data[N29], Data[N13], Data[N32], Data[N34], Data[N9], Data[N33], Data[N15], Data[N11], Data[N17], Data[N36], Data[N31], Data[N14], Data[N18], Data[N19], Data[N16], Data[N35], Data[N37]

The symbolic expression is:
((((((((((((((((((((((((((((((((!(((((!(IN4)) & (!(IN2))) & (!(IN22))) & (!(IN3))) & (!(IN21)))) | IN1) & ((!((((IN4 & (!(IN2))) & (!(IN22))) & (!(IN3))) & (!(IN21)))) | IN5)) & ((!(((((!(IN4)) & IN2) & (!(IN22))) & (!(IN3))) & (!(IN21)))) | IN20)) & ((!((((IN4 & IN2) & (!(IN22))) & (!(IN3))) & (!(IN21)))) | IN7)) & ((!(((((!(IN4)) & (!(IN2))) & IN22) & (!(IN3))) & (!(IN21)))) | IN6)) & ((!((((IN4 & (!(IN2))) & IN22) & (!(IN3))) & (!(IN21)))) | IN8)) & ((!(((((!(IN4)) & IN2) & IN22) & (!(IN3))) & (!(IN21)))) | IN23)) & ((!((((IN4 & IN2) & IN22) & (!(IN3))) & (!(IN21)))) | IN10)) & ((!(((((!(IN4)) & (!(IN2))) & (!(IN22))) & IN3) & (!(IN21)))) | IN26)) & ((!((((IN4 & (!(IN2))) & (!(IN22))) & IN3) & (!(IN21)))) | IN28)) & ((!(((((!(IN4)) & IN2) & (!(IN22))) & IN3) & (!(IN21)))) | IN25)) & ((!((((IN4 & IN2) & (!(IN22))) & IN3) & (!(IN21)))) | IN27)) & ((!(((((!(IN4)) & (!(IN2))) & IN22) & IN3) & (!(IN21)))) | IN12)) & ((!((((IN4 & (!(IN2))) & IN22) & IN3) & (!(IN21)))) | IN30)) & ((!(((((!(IN4)) & IN2) & IN22) & IN3) & (!(IN21)))) | IN24)) & ((!((((IN4 & IN2) & IN22) & IN3) & (!(IN21)))) | IN29)) & ((!(((((!(IN4)) & (!(IN2))) & (!(IN22))) & (!(IN3))) & IN21)) | IN13)) & ((!((((IN4 & (!(IN2))) & (!(IN22))) & (!(IN3))) & IN21)) | IN32)) & ((!(((((!(IN4)) & IN2) & (!(IN22))) & (!(IN3))) & IN21)) | IN34)) & ((!((((IN4 & IN2) & (!(IN22))) & (!(IN3))) & IN21)) | IN9)) & ((!(((((!(IN4)) & (!(IN2))) & IN22) & (!(IN3))) & IN21)) | IN33)) & ((!((((IN4 & (!(IN2))) & IN22) & (!(IN3))) & IN21)) | IN15)) & ((!(((((!(IN4)) & IN2) & IN22) & (!(IN3))) & IN21)) | IN11)) & ((!((((IN4 & IN2) & IN22) & (!(IN3))) & IN21)) | IN17)) & ((!(((((!(IN4)) & (!(IN2))) & (!(IN22))) & IN3) & IN21)) | IN36)) & ((!((((IN4 & (!(IN2))) & (!(IN22))) & IN3) & IN21)) | IN31)) & ((!(((((!(IN4)) & IN2) & (!(IN22))) & IN3) & IN21)) | IN14)) & ((!((((IN4 & IN2) & (!(IN22))) & IN3) & IN21)) | IN18)) & ((!(((((!(IN4)) & (!(IN2))) & IN22) & IN3) & IN21)) | IN19)) & ((!((((IN4 & (!(IN2))) & IN22) & IN3) & IN21)) | IN16)) & ((!(((((!(IN4)) & IN2) & IN22) & IN3) & IN21)) | IN35)) & ((!((((IN4 & IN2) & IN22) & IN3) & IN21)) | IN37)

*)

FUNCTION_BLOCK F_CollectInput
  VAR_IN_OUT
      Data : ARRAY[1..40] OF BOOL;
  END_VAR
  VAR_INPUT
      TICK  : BOOL := 0;
      IN1   : BOOL := 0;
      IN2   : BOOL := 0;
      IN3   : BOOL := 0;
      IN4   : BOOL := 0;
      IN5   : BOOL := 0;
      RESET : BOOL := FALSE;
  END_VAR
  VAR_OUTPUT
      Finished : BOOL;
  END_VAR
  VAR
      j    : USINT := 1;
      tock : BOOL  := 0;
  END_VAR
  IF NOT RESET AND tock = NOT TICK THEN
      Data[j]   := IN1;
      Data[j+1] := IN2;
      Data[j+2] := IN3;
      Data[j+3] := IN4;
      Data[j+4] := IN5;
      j := j + 5;
      tock := TICK;
  ELSE
      j := 1;
      tock := 0;
  END_IF;
  Finished := (j > 40);
END_FUNCTION_BLOCK

PROGRAM Boiler
  VAR
    Data  : ARRAY[1..40] OF BOOL;
    Ready : BOOL;
    CollectInput : F_CollectInput;
  END_VAR
  VAR
    TICK     AT %IX1.0 : BOOL;
    IN1      AT %IX0.3 : BOOL;
    IN2      AT %IX0.4 : BOOL;
    IN3      AT %IX0.5 : BOOL;
    IN4      AT %IX0.6 : BOOL;
    IN5      AT %IX0.7 : BOOL;
    OutReady AT %QX0.0 : BOOL := FALSE;
    FeedNext AT %QX0.1 : BOOL := FALSE;
    Out      AT %QX0.2 : BOOL;
  END_VAR
  CollectInput(TICK:=TICK, IN1:=IN1, IN2:=IN2, IN3:=IN3, IN4:=IN4, IN5:=IN5);
  Ready := CollectInput.Finished;
  FeedNext := 1;
  IF Ready THEN
    Out := (((((((((((((((((((((((((((((((((NOT (((((NOT Data[4]) AND (NOT Data[2])) AND (NOT Data[22])) AND (NOT Data[3])) AND (NOT Data[21]))) OR Data[1]) AND ((NOT ((((Data[4] AND (NOT Data[2])) AND (NOT Data[22])) AND (NOT Data[3])) AND (NOT Data[21]))) OR Data[5])) AND ((NOT (((((NOT Data[4]) AND Data[2]) AND (NOT Data[22])) AND (NOT Data[3])) AND (NOT Data[21]))) OR Data[20])) AND ((NOT ((((Data[4] AND Data[2]) AND (NOT Data[22])) AND (NOT Data[3])) AND (NOT Data[21]))) OR Data[7])) AND ((NOT (((((NOT Data[4]) AND (NOT Data[2])) AND Data[22]) AND (NOT Data[3])) AND (NOT Data[21]))) OR Data[6])) AND ((NOT ((((Data[4] AND (NOT Data[2])) AND Data[22]) AND (NOT Data[3])) AND (NOT Data[21]))) OR Data[8])) AND ((NOT (((((NOT Data[4]) AND Data[2]) AND Data[22]) AND (NOT Data[3])) AND (NOT Data[21]))) OR Data[23])) AND ((NOT ((((Data[4] AND Data[2]) AND Data[22]) AND (NOT Data[3])) AND (NOT Data[21]))) OR Data[10])) AND ((NOT (((((NOT Data[4]) AND (NOT Data[2])) AND (NOT Data[22])) AND Data[3]) AND (NOT Data[21]))) OR Data[26])) AND ((NOT ((((Data[4] AND (NOT Data[2])) AND (NOT Data[22])) AND Data[3]) AND (NOT Data[21]))) OR Data[28])) AND ((NOT (((((NOT Data[4]) AND Data[2]) AND (NOT Data[22])) AND Data[3]) AND (NOT Data[21]))) OR Data[25])) AND ((NOT ((((Data[4] AND Data[2]) AND (NOT Data[22])) AND Data[3]) AND (NOT Data[21]))) OR Data[27])) AND ((NOT (((((NOT Data[4]) AND (NOT Data[2])) AND Data[22]) AND Data[3]) AND (NOT Data[21]))) OR Data[12])) AND ((NOT ((((Data[4] AND (NOT Data[2])) AND Data[22]) AND Data[3]) AND (NOT Data[21]))) OR Data[30])) AND ((NOT (((((NOT Data[4]) AND Data[2]) AND Data[22]) AND Data[3]) AND (NOT Data[21]))) OR Data[24])) AND ((NOT ((((Data[4] AND Data[2]) AND Data[22]) AND Data[3]) AND (NOT Data[21]))) OR Data[29])) AND ((NOT (((((NOT Data[4]) AND (NOT Data[2])) AND (NOT Data[22])) AND (NOT Data[3])) AND Data[21])) OR Data[13])) AND ((NOT ((((Data[4] AND (NOT Data[2])) AND (NOT Data[22])) AND (NOT Data[3])) AND Data[21])) OR Data[32])) AND ((NOT (((((NOT Data[4]) AND Data[2]) AND (NOT Data[22])) AND (NOT Data[3])) AND Data[21])) OR Data[34])) AND ((NOT ((((Data[4] AND Data[2]) AND (NOT Data[22])) AND (NOT Data[3])) AND Data[21])) OR Data[9])) AND ((NOT (((((NOT Data[4]) AND (NOT Data[2])) AND Data[22]) AND (NOT Data[3])) AND Data[21])) OR Data[33])) AND ((NOT ((((Data[4] AND (NOT Data[2])) AND Data[22]) AND (NOT Data[3])) AND Data[21])) OR Data[15])) AND ((NOT (((((NOT Data[4]) AND Data[2]) AND Data[22]) AND (NOT Data[3])) AND Data[21])) OR Data[11])) AND ((NOT ((((Data[4] AND Data[2]) AND Data[22]) AND (NOT Data[3])) AND Data[21])) OR Data[17])) AND ((NOT (((((NOT Data[4]) AND (NOT Data[2])) AND (NOT Data[22])) AND Data[3]) AND Data[21])) OR Data[36])) AND ((NOT ((((Data[4] AND (NOT Data[2])) AND (NOT Data[22])) AND Data[3]) AND Data[21])) OR Data[31])) AND ((NOT (((((NOT Data[4]) AND Data[2]) AND (NOT Data[22])) AND Data[3]) AND Data[21])) OR Data[14])) AND ((NOT ((((Data[4] AND Data[2]) AND (NOT Data[22])) AND Data[3]) AND Data[21])) OR Data[18])) AND ((NOT (((((NOT Data[4]) AND (NOT Data[2])) AND Data[22]) AND Data[3]) AND Data[21])) OR Data[19])) AND ((NOT ((((Data[4] AND (NOT Data[2])) AND Data[22]) AND Data[3]) AND Data[21])) OR Data[16])) AND ((NOT (((((NOT Data[4]) AND Data[2]) AND Data[22]) AND Data[3]) AND Data[21])) OR Data[35])) AND ((NOT ((((Data[4] AND Data[2]) AND Data[22]) AND Data[3]) AND Data[21])) OR Data[37]));
    OutReady := 1;
    CollectInput(RESET:=TRUE);
  END_IF;
END_PROGRAM

CONFIGURATION Config0
  RESOURCE Res0 ON PLC
    TASK task0(INTERVAL := T#20ms,PRIORITY := 0);
    PROGRAM instance0 WITH task0 : Boiler;
  END_RESOURCE
END_CONFIGURATION

(* ---- 5-MUX_zebus-blank-faddy.st ---- *)
(*
This code implements a shuffled multiplexer with 5 control bits.
The control bits are: Data[N1], Data[N2], Data[N3], Data[N4], Data[N20]
The input bits are: Data[N5], Data[N8], Data[N6], Data[N23], Data[N22], Data[N21], Data[N9], Data[N24], Data[N7], Data[N25], Data[N26], Data[N30], Data[N28], Data[N27], Data[N10], Data[N11], Data[N14], Data[N12], Data[N31], Data[N32], Data[N29], Data[N13], Data[N35], Data[N16], Data[N19], Data[N17], Data[N15], Data[N33], Data[N18], Data[N37], Data[N34], Data[N36]

The symbolic expression is:
((((((((((((((((((((((((((((((((!(((((!(IN1)) & (!(IN2))) & (!(IN3))) & (!(IN4))) & (!(IN20)))) | IN5) & ((!((((IN1 & (!(IN2))) & (!(IN3))) & (!(IN4))) & (!(IN20)))) | IN8)) & ((!(((((!(IN1)) & IN2) & (!(IN3))) & (!(IN4))) & (!(IN20)))) | IN6)) & ((!((((IN1 & IN2) & (!(IN3))) & (!(IN4))) & (!(IN20)))) | IN23)) & ((!(((((!(IN1)) & (!(IN2))) & IN3) & (!(IN4))) & (!(IN20)))) | IN22)) & ((!((((IN1 & (!(IN2))) & IN3) & (!(IN4))) & (!(IN20)))) | IN21)) & ((!(((((!(IN1)) & IN2) & IN3) & (!(IN4))) & (!(IN20)))) | IN9)) & ((!((((IN1 & IN2) & IN3) & (!(IN4))) & (!(IN20)))) | IN24)) & ((!(((((!(IN1)) & (!(IN2))) & (!(IN3))) & IN4) & (!(IN20)))) | IN7)) & ((!((((IN1 & (!(IN2))) & (!(IN3))) & IN4) & (!(IN20)))) | IN25)) & ((!(((((!(IN1)) & IN2) & (!(IN3))) & IN4) & (!(IN20)))) | IN26)) & ((!((((IN1 & IN2) & (!(IN3))) & IN4) & (!(IN20)))) | IN30)) & ((!(((((!(IN1)) & (!(IN2))) & IN3) & IN4) & (!(IN20)))) | IN28)) & ((!((((IN1 & (!(IN2))) & IN3) & IN4) & (!(IN20)))) | IN27)) & ((!(((((!(IN1)) & IN2) & IN3) & IN4) & (!(IN20)))) | IN10)) & ((!((((IN1 & IN2) & IN3) & IN4) & (!(IN20)))) | IN11)) & ((!(((((!(IN1)) & (!(IN2))) & (!(IN3))) & (!(IN4))) & IN20)) | IN14)) & ((!((((IN1 & (!(IN2))) & (!(IN3))) & (!(IN4))) & IN20)) | IN12)) & ((!(((((!(IN1)) & IN2) & (!(IN3))) & (!(IN4))) & IN20)) | IN31)) & ((!((((IN1 & IN2) & (!(IN3))) & (!(IN4))) & IN20)) | IN32)) & ((!(((((!(IN1)) & (!(IN2))) & IN3) & (!(IN4))) & IN20)) | IN29)) & ((!((((IN1 & (!(IN2))) & IN3) & (!(IN4))) & IN20)) | IN13)) & ((!(((((!(IN1)) & IN2) & IN3) & (!(IN4))) & IN20)) | IN35)) & ((!((((IN1 & IN2) & IN3) & (!(IN4))) & IN20)) | IN16)) & ((!(((((!(IN1)) & (!(IN2))) & (!(IN3))) & IN4) & IN20)) | IN19)) & ((!((((IN1 & (!(IN2))) & (!(IN3))) & IN4) & IN20)) | IN17)) & ((!(((((!(IN1)) & IN2) & (!(IN3))) & IN4) & IN20)) | IN15)) & ((!((((IN1 & IN2) & (!(IN3))) & IN4) & IN20)) | IN33)) & ((!(((((!(IN1)) & (!(IN2))) & IN3) & IN4) & IN20)) | IN18)) & ((!((((IN1 & (!(IN2))) & IN3) & IN4) & IN20)) | IN37)) & ((!(((((!(IN1)) & IN2) & IN3) & IN4) & IN20)) | IN34)) & ((!((((IN1 & IN2) & IN3) & IN4) & IN20)) | IN36)

*)

FUNCTION_BLOCK F_CollectInput
  VAR_IN_OUT
      Data : ARRAY[1..40] OF BOOL;
  END_VAR
  VAR_INPUT
      TICK  : BOOL := 0;
      IN1   : BOOL := 0;
      IN2   : BOOL := 0;
      IN3   : BOOL := 0;
      IN4   : BOOL := 0;
      IN5   : BOOL := 0;
      RESET : BOOL := FALSE;
  END_VAR
  VAR_OUTPUT
      Finished : BOOL;
  END_VAR
  VAR
      j    : USINT := 1;
      tock : BOOL  := 0;
  END_VAR
  IF NOT RESET AND tock = NOT TICK THEN
      Data[j]   := IN1;
      Data[j+1] := IN2;
      Data[j+2] := IN3;
      Data[j+3] := IN4;
      Data[j+4] := IN5;
      j := j + 5;
      tock := TICK;
  ELSE
      j := 1;
      tock := 0;
  END_IF;
  Finished := (j > 40);
END_FUNCTION_BLOCK

PROGRAM Boiler
  VAR
    Data  : ARRAY[1..40] OF BOOL;
    Ready : BOOL;
    CollectInput : F_CollectInput;
  END_VAR
  VAR
    TICK     AT %IX1.0 : BOOL;
    IN1      AT %IX0.3 : BOOL;
    IN2      AT %IX0.4 : BOOL;
    IN3      AT %IX0.5 : BOOL;
    IN4      AT %IX0.6 : BOOL;
    IN5      AT %IX0.7 : BOOL;
    OutReady AT %QX0.0 : BOOL := FALSE;
    FeedNext AT %QX0.1 : BOOL := FALSE;
    Out      AT %QX0.2 : BOOL;
  END_VAR
  CollectInput(TICK:=TICK, IN1:=IN1, IN2:=IN2, IN3:=IN3, IN4:=IN4, IN5:=IN5);
  Ready := CollectInput.Finished;
  FeedNext := 1;
  IF Ready THEN
    Out := (((((((((((((((((((((((((((((((((NOT (((((NOT Data[1]) AND (NOT Data[2])) AND (NOT Data[3])) AND (NOT Data[4])) AND (NOT Data[20]))) OR Data[5]) AND ((NOT ((((Data[1] AND (NOT Data[2])) AND (NOT Data[3])) AND (NOT Data[4])) AND (NOT Data[20]))) OR Data[8])) AND ((NOT (((((NOT Data[1]) AND Data[2]) AND (NOT Data[3])) AND (NOT Data[4])) AND (NOT Data[20]))) OR Data[6])) AND ((NOT ((((Data[1] AND Data[2]) AND (NOT Data[3])) AND (NOT Data[4])) AND (NOT Data[20]))) OR Data[23])) AND ((NOT (((((NOT Data[1]) AND (NOT Data[2])) AND Data[3]) AND (NOT Data[4])) AND (NOT Data[20]))) OR Data[22])) AND ((NOT ((((Data[1] AND (NOT Data[2])) AND Data[3]) AND (NOT Data[4])) AND (NOT Data[20]))) OR Data[21])) AND ((NOT (((((NOT Data[1]) AND Data[2]) AND Data[3]) AND (NOT Data[4])) AND (NOT Data[20]))) OR Data[9])) AND ((NOT ((((Data[1] AND Data[2]) AND Data[3]) AND (NOT Data[4])) AND (NOT Data[20]))) OR Data[24])) AND ((NOT (((((NOT Data[1]) AND (NOT Data[2])) AND (NOT Data[3])) AND Data[4]) AND (NOT Data[20]))) OR Data[7])) AND ((NOT ((((Data[1] AND (NOT Data[2])) AND (NOT Data[3])) AND Data[4]) AND (NOT Data[20]))) OR Data[25])) AND ((NOT (((((NOT Data[1]) AND Data[2]) AND (NOT Data[3])) AND Data[4]) AND (NOT Data[20]))) OR Data[26])) AND ((NOT ((((Data[1] AND Data[2]) AND (NOT Data[3])) AND Data[4]) AND (NOT Data[20]))) OR Data[30])) AND ((NOT (((((NOT Data[1]) AND (NOT Data[2])) AND Data[3]) AND Data[4]) AND (NOT Data[20]))) OR Data[28])) AND ((NOT ((((Data[1] AND (NOT Data[2])) AND Data[3]) AND Data[4]) AND (NOT Data[20]))) OR Data[27])) AND ((NOT (((((NOT Data[1]) AND Data[2]) AND Data[3]) AND Data[4]) AND (NOT Data[20]))) OR Data[10])) AND ((NOT ((((Data[1] AND Data[2]) AND Data[3]) AND Data[4]) AND (NOT Data[20]))) OR Data[11])) AND ((NOT (((((NOT Data[1]) AND (NOT Data[2])) AND (NOT Data[3])) AND (NOT Data[4])) AND Data[20])) OR Data[14])) AND ((NOT ((((Data[1] AND (NOT Data[2])) AND (NOT Data[3])) AND (NOT Data[4])) AND Data[20])) OR Data[12])) AND ((NOT (((((NOT Data[1]) AND Data[2]) AND (NOT Data[3])) AND (NOT Data[4])) AND Data[20])) OR Data[31])) AND ((NOT ((((Data[1] AND Data[2]) AND (NOT Data[3])) AND (NOT Data[4])) AND Data[20])) OR Data[32])) AND ((NOT (((((NOT Data[1]) AND (NOT Data[2])) AND Data[3]) AND (NOT Data[4])) AND Data[20])) OR Data[29])) AND ((NOT ((((Data[1] AND (NOT Data[2])) AND Data[3]) AND (NOT Data[4])) AND Data[20])) OR Data[13])) AND ((NOT (((((NOT Data[1]) AND Data[2]) AND Data[3]) AND (NOT Data[4])) AND Data[20])) OR Data[35])) AND ((NOT ((((Data[1] AND Data[2]) AND Data[3]) AND (NOT Data[4])) AND Data[20])) OR Data[16])) AND ((NOT (((((NOT Data[1]) AND (NOT Data[2])) AND (NOT Data[3])) AND Data[4]) AND Data[20])) OR Data[19])) AND ((NOT ((((Data[1] AND (NOT Data[2])) AND (NOT Data[3])) AND Data[4]) AND Data[20])) OR Data[17])) AND ((NOT (((((NOT Data[1]) AND Data[2]) AND (NOT Data[3])) AND Data[4]) AND Data[20])) OR Data[15])) AND ((NOT ((((Data[1] AND Data[2]) AND (NOT Data[3])) AND Data[4]) AND Data[20])) OR Data[33])) AND ((NOT (((((NOT Data[1]) AND (NOT Data[2])) AND Data[3]) AND Data[4]) AND Data[20])) OR Data[18])) AND ((NOT ((((Data[1] AND (NOT Data[2])) AND Data[3]) AND Data[4]) AND Data[20])) OR Data[37])) AND ((NOT (((((NOT Data[1]) AND Data[2]) AND Data[3]) AND Data[4]) AND Data[20])) OR Data[34])) AND ((NOT ((((Data[1] AND Data[2]) AND Data[3]) AND Data[4]) AND Data[20])) OR Data[36]));
    OutReady := 1;
    CollectInput(RESET:=TRUE);
  END_IF;
END_PROGRAM

CONFIGURATION Config0
  RESOURCE Res0 ON PLC
    TASK task0(INTERVAL := T#20ms,PRIORITY := 0);
    PROGRAM instance0 WITH task0 : Boiler;
  END_RESOURCE
END_CONFIGURATION

(* ---- 5-MUX_zonal-brink-sassy.st ---- *)
(*
This code implements a shuffled multiplexer with 5 control bits.
The control bits are: Data[N1], Data[N2], Data[N25], Data[N23], Data[N22]
The input bits are: Data[N20], Data[N3], Data[N21], Data[N8], Data[N24], Data[N26], Data[N4], Data[N10], Data[N27], Data[N6], Data[N28], Data[N31], Data[N32], Data[N29], Data[N30], Data[N11], Data[N13], Data[N7], Data[N9], Data[N35], Data[N36], Data[N16], Data[N34], Data[N5], Data[N37], Data[N14], Data[N15], Data[N19], Data[N33], Data[N12], Data[N17], Data[N18]

The symbolic expression is:
((((((((((((((((((((((((((((((((!(((((!(IN1)) & (!(IN2))) & (!(IN25))) & (!(IN23))) & (!(IN22)))) | IN20) & ((!((((IN1 & (!(IN2))) & (!(IN25))) & (!(IN23))) & (!(IN22)))) | IN3)) & ((!(((((!(IN1)) & IN2) & (!(IN25))) & (!(IN23))) & (!(IN22)))) | IN21)) & ((!((((IN1 & IN2) & (!(IN25))) & (!(IN23))) & (!(IN22)))) | IN8)) & ((!(((((!(IN1)) & (!(IN2))) & IN25) & (!(IN23))) & (!(IN22)))) | IN24)) & ((!((((IN1 & (!(IN2))) & IN25) & (!(IN23))) & (!(IN22)))) | IN26)) & ((!(((((!(IN1)) & IN2) & IN25) & (!(IN23))) & (!(IN22)))) | IN4)) & ((!((((IN1 & IN2) & IN25) & (!(IN23))) & (!(IN22)))) | IN10)) & ((!(((((!(IN1)) & (!(IN2))) & (!(IN25))) & IN23) & (!(IN22)))) | IN27)) & ((!((((IN1 & (!(IN2))) & (!(IN25))) & IN23) & (!(IN22)))) | IN6)) & ((!(((((!(IN1)) & IN2) & (!(IN25))) & IN23) & (!(IN22)))) | IN28)) & ((!((((IN1 & IN2) & (!(IN25))) & IN23) & (!(IN22)))) | IN31)) & ((!(((((!(IN1)) & (!(IN2))) & IN25) & IN23) & (!(IN22)))) | IN32)) & ((!((((IN1 & (!(IN2))) & IN25) & IN23) & (!(IN22)))) | IN29)) & ((!(((((!(IN1)) & IN2) & IN25) & IN23) & (!(IN22)))) | IN30)) & ((!((((IN1 & IN2) & IN25) & IN23) & (!(IN22)))) | IN11)) & ((!(((((!(IN1)) & (!(IN2))) & (!(IN25))) & (!(IN23))) & IN22)) | IN13)) & ((!((((IN1 & (!(IN2))) & (!(IN25))) & (!(IN23))) & IN22)) | IN7)) & ((!(((((!(IN1)) & IN2) & (!(IN25))) & (!(IN23))) & IN22)) | IN9)) & ((!((((IN1 & IN2) & (!(IN25))) & (!(IN23))) & IN22)) | IN35)) & ((!(((((!(IN1)) & (!(IN2))) & IN25) & (!(IN23))) & IN22)) | IN36)) & ((!((((IN1 & (!(IN2))) & IN25) & (!(IN23))) & IN22)) | IN16)) & ((!(((((!(IN1)) & IN2) & IN25) & (!(IN23))) & IN22)) | IN34)) & ((!((((IN1 & IN2) & IN25) & (!(IN23))) & IN22)) | IN5)) & ((!(((((!(IN1)) & (!(IN2))) & (!(IN25))) & IN23) & IN22)) | IN37)) & ((!((((IN1 & (!(IN2))) & (!(IN25))) & IN23) & IN22)) | IN14)) & ((!(((((!(IN1)) & IN2) & (!(IN25))) & IN23) & IN22)) | IN15)) & ((!((((IN1 & IN2) & (!(IN25))) & IN23) & IN22)) | IN19)) & ((!(((((!(IN1)) & (!(IN2))) & IN25) & IN23) & IN22)) | IN33)) & ((!((((IN1 & (!(IN2))) & IN25) & IN23) & IN22)) | IN12)) & ((!(((((!(IN1)) & IN2) & IN25) & IN23) & IN22)) | IN17)) & ((!((((IN1 & IN2) & IN25) & IN23) & IN22)) | IN18)

*)

FUNCTION_BLOCK F_CollectInput
  VAR_IN_OUT
      Data : ARRAY[1..40] OF BOOL;
  END_VAR
  VAR_INPUT
      TICK  : BOOL := 0;
      IN1   : BOOL := 0;
      IN2   : BOOL := 0;
      IN3   : BOOL := 0;
      IN4   : BOOL := 0;
      IN5   : BOOL := 0;
      RESET : BOOL := FALSE;
  END_VAR
  VAR_OUTPUT
      Finished : BOOL;
  END_VAR
  VAR
      j    : USINT := 1;
      tock : BOOL  := 0;
  END_VAR
  IF NOT RESET AND tock = NOT TICK THEN
      Data[j]   := IN1;
      Data[j+1] := IN2;
      Data[j+2] := IN3;
      Data[j+3] := IN4;
      Data[j+4] := IN5;
      j := j + 5;
      tock := TICK;
  ELSE
      j := 1;
      tock := 0;
  END_IF;
  Finished := (j > 40);
END_FUNCTION_BLOCK

PROGRAM Boiler
  VAR
    Data  : ARRAY[1..40] OF BOOL;
    Ready : BOOL;
    CollectInput : F_CollectInput;
  END_VAR
  VAR
    TICK     AT %IX1.0 : BOOL;
    IN1      AT %IX0.3 : BOOL;
    IN2      AT %IX0.4 : BOOL;
    IN3      AT %IX0.5 : BOOL;
    IN4      AT %IX0.6 : BOOL;
    IN5      AT %IX0.7 : BOOL;
    OutReady AT %QX0.0 : BOOL := FALSE;
    FeedNext AT %QX0.1 : BOOL := FALSE;
    Out      AT %QX0.2 : BOOL;
  END_VAR
  CollectInput(TICK:=TICK, IN1:=IN1, IN2:=IN2, IN3:=IN3, IN4:=IN4, IN5:=IN5);
  Ready := CollectInput.Finished;
  FeedNext := 1;
  IF Ready THEN
    Out := (((((((((((((((((((((((((((((((((NOT (((((NOT Data[1]) AND (NOT Data[2])) AND (NOT Data[25])) AND (NOT Data[23])) AND (NOT Data[22]))) OR Data[20]) AND ((NOT ((((Data[1] AND (NOT Data[2])) AND (NOT Data[25])) AND (NOT Data[23])) AND (NOT Data[22]))) OR Data[3])) AND ((NOT (((((NOT Data[1]) AND Data[2]) AND (NOT Data[25])) AND (NOT Data[23])) AND (NOT Data[22]))) OR Data[21])) AND ((NOT ((((Data[1] AND Data[2]) AND (NOT Data[25])) AND (NOT Data[23])) AND (NOT Data[22]))) OR Data[8])) AND ((NOT (((((NOT Data[1]) AND (NOT Data[2])) AND Data[25]) AND (NOT Data[23])) AND (NOT Data[22]))) OR Data[24])) AND ((NOT ((((Data[1] AND (NOT Data[2])) AND Data[25]) AND (NOT Data[23])) AND (NOT Data[22]))) OR Data[26])) AND ((NOT (((((NOT Data[1]) AND Data[2]) AND Data[25]) AND (NOT Data[23])) AND (NOT Data[22]))) OR Data[4])) AND ((NOT ((((Data[1] AND Data[2]) AND Data[25]) AND (NOT Data[23])) AND (NOT Data[22]))) OR Data[10])) AND ((NOT (((((NOT Data[1]) AND (NOT Data[2])) AND (NOT Data[25])) AND Data[23]) AND (NOT Data[22]))) OR Data[27])) AND ((NOT ((((Data[1] AND (NOT Data[2])) AND (NOT Data[25])) AND Data[23]) AND (NOT Data[22]))) OR Data[6])) AND ((NOT (((((NOT Data[1]) AND Data[2]) AND (NOT Data[25])) AND Data[23]) AND (NOT Data[22]))) OR Data[28])) AND ((NOT ((((Data[1] AND Data[2]) AND (NOT Data[25])) AND Data[23]) AND (NOT Data[22]))) OR Data[31])) AND ((NOT (((((NOT Data[1]) AND (NOT Data[2])) AND Data[25]) AND Data[23]) AND (NOT Data[22]))) OR Data[32])) AND ((NOT ((((Data[1] AND (NOT Data[2])) AND Data[25]) AND Data[23]) AND (NOT Data[22]))) OR Data[29])) AND ((NOT (((((NOT Data[1]) AND Data[2]) AND Data[25]) AND Data[23]) AND (NOT Data[22]))) OR Data[30])) AND ((NOT ((((Data[1] AND Data[2]) AND Data[25]) AND Data[23]) AND (NOT Data[22]))) OR Data[11])) AND ((NOT (((((NOT Data[1]) AND (NOT Data[2])) AND (NOT Data[25])) AND (NOT Data[23])) AND Data[22])) OR Data[13])) AND ((NOT ((((Data[1] AND (NOT Data[2])) AND (NOT Data[25])) AND (NOT Data[23])) AND Data[22])) OR Data[7])) AND ((NOT (((((NOT Data[1]) AND Data[2]) AND (NOT Data[25])) AND (NOT Data[23])) AND Data[22])) OR Data[9])) AND ((NOT ((((Data[1] AND Data[2]) AND (NOT Data[25])) AND (NOT Data[23])) AND Data[22])) OR Data[35])) AND ((NOT (((((NOT Data[1]) AND (NOT Data[2])) AND Data[25]) AND (NOT Data[23])) AND Data[22])) OR Data[36])) AND ((NOT ((((Data[1] AND (NOT Data[2])) AND Data[25]) AND (NOT Data[23])) AND Data[22])) OR Data[16])) AND ((NOT (((((NOT Data[1]) AND Data[2]) AND Data[25]) AND (NOT Data[23])) AND Data[22])) OR Data[34])) AND ((NOT ((((Data[1] AND Data[2]) AND Data[25]) AND (NOT Data[23])) AND Data[22])) OR Data[5])) AND ((NOT (((((NOT Data[1]) AND (NOT Data[2])) AND (NOT Data[25])) AND Data[23]) AND Data[22])) OR Data[37])) AND ((NOT ((((Data[1] AND (NOT Data[2])) AND (NOT Data[25])) AND Data[23]) AND Data[22])) OR Data[14])) AND ((NOT (((((NOT Data[1]) AND Data[2]) AND (NOT Data[25])) AND Data[23]) AND Data[22])) OR Data[15])) AND ((NOT ((((Data[1] AND Data[2]) AND (NOT Data[25])) AND Data[23]) AND Data[22])) OR Data[19])) AND ((NOT (((((NOT Data[1]) AND (NOT Data[2])) AND Data[25]) AND Data[23]) AND Data[22])) OR Data[33])) AND ((NOT ((((Data[1] AND (NOT Data[2])) AND Data[25]) AND Data[23]) AND Data[22])) OR Data[12])) AND ((NOT (((((NOT Data[1]) AND Data[2]) AND Data[25]) AND Data[23]) AND Data[22])) OR Data[17])) AND ((NOT ((((Data[1] AND Data[2]) AND Data[25]) AND Data[23]) AND Data[22])) OR Data[18]));
    OutReady := 1;
    CollectInput(RESET:=TRUE);
  END_IF;
END_PROGRAM

CONFIGURATION Config0
  RESOURCE Res0 ON PLC
    TASK task0(INTERVAL := T#20ms,PRIORITY := 0);
    PROGRAM instance0 WITH task0 : Boiler;
  END_RESOURCE
END_CONFIGURATION

(* ---- RND-EXPR_8var-dicey-verbs-seeds.st ---- *)
FUNCTION_BLOCK F_CollectInput
  VAR_IN_OUT
      Data : ARRAY[1..10] OF BOOL;
  END_VAR
  VAR_INPUT
      TICK  : BOOL := 0;
      IN1   : BOOL := 0;
      IN2   : BOOL := 0;
      IN3   : BOOL := 0;
      IN4   : BOOL := 0;
      IN5   : BOOL := 0;
      RESET : BOOL := FALSE;
  END_VAR
  VAR_OUTPUT
      Finished : BOOL;
  END_VAR
  VAR
      j    : USINT := 1;
      tock : BOOL  := 0;
  END_VAR
  IF NOT RESET AND tock = NOT TICK THEN
      Data[j]   := IN1;
      Data[j+1] := IN2;
      Data[j+2] := IN3;
      Data[j+3] := IN4;
      Data[j+4] := IN5;
      j := j + 5;
      tock := TICK;
  ELSE
      j := 1;
      tock := 0;
  END_IF;
  Finished := (j > 10);
END_FUNCTION_BLOCK

PROGRAM Boiler
  VAR
    Data  : ARRAY[1..10] OF BOOL;
    Ready : BOOL;
    CollectInput : F_CollectInput;
  END_VAR
  VAR
    TICK     AT %IX1.0 : BOOL;
    IN1      AT %IX0.3 : BOOL;
    IN2      AT %IX0.4 : BOOL;
    IN3      AT %IX0.5 : BOOL;
    IN4      AT %IX0.6 : BOOL;
    IN5      AT %IX0.7 : BOOL;
    OutReady AT %QX0.0 : BOOL := FALSE;
    FeedNext AT %QX0.1 : BOOL := FALSE;
    Out      AT %QX0.2 : BOOL;
  END_VAR
  CollectInput(TICK:=TICK, IN1:=IN1, IN2:=IN2, IN3:=IN3, IN4:=IN4, IN5:=IN5);
  Ready := CollectInput.Finished;
  FeedNext := 1;
  IF Ready THEN
    Out := ((NOT ((((NOT D[3]) OR ((NOT (NOT D[4])) AND D[8])) OR TRUE) AND ((NOT D[4]) AND ((((NOT ((D[4] OR ((NOT (NOT D[6])) OR ((D[8] OR D[2]) AND (NOT D[2])))) AND (((TRUE OR (TRUE OR FALSE)) OR ((D[5] AND D[5]) OR (TRUE AND D[1]))) AND ((NOT (NOT D[8])) AND ((D[2] AND D[2]) OR (D[2] OR FALSE)))))) AND (NOT (((((NOT D[4]) OR (NOT D[7])) AND ((NOT D[2]) OR (NOT D[2]))) AND TRUE) AND TRUE))) AND (((NOT ((D[2] AND (D[6] OR (D[3] AND D[8]))) AND (NOT D[6]))) AND ((NOT D[8]) OR (D[8] AND (NOT (NOT (D[8] AND D[2])))))) AND ((((NOT ((D[5] OR D[8]) AND (D[6] OR D[3]))) OR (((NOT D[8]) OR D[5]) AND ((D[3] AND D[3]) OR (NOT D[2])))) OR (NOT D[2])) OR (((((D[7] OR D[6]) AND (NOT D[1])) AND ((NOT D[6]) AND (D[3] AND D[6]))) AND (((TRUE OR D[8]) AND (D[4] AND D[6])) OR ((D[7] OR D[1]) AND (D[6] AND D[7])))) OR (NOT ((D[2] OR (D[4] OR FALSE)) OR ((NOT D[3]) OR (TRUE AND D[7])))))))) OR ((NOT ((D[1] OR (((NOT (D[2] OR D[6])) OR D[7]) AND ((NOT (D[8] OR D[4])) OR ((NOT D[7]) OR (D[5] AND D[1]))))) OR D[5])) OR (((NOT ((((TRUE OR TRUE) OR D[5]) AND (D[3] AND (NOT D[4]))) AND (((D[1] AND D[1]) AND (D[6] OR D[1])) AND ((D[7] AND D[2]) OR (D[8] AND FALSE))))) OR ((NOT ((NOT (D[4] AND D[2])) AND (NOT (NOT D[4])))) AND ((NOT ((D[2] AND D[8]) AND (D[6] AND D[4]))) OR D[2]))) AND ((((D[6] OR (NOT (D[6] AND D[3]))) AND (((NOT D[3]) OR D[7]) OR ((D[6] OR D[6]) AND (NOT D[5])))) AND TRUE) OR (((NOT D[7]) OR FALSE) OR (NOT ((NOT (D[8] OR D[4])) AND (NOT (D[4] OR FALSE)))))))))))) OR D[7]);
    OutReady := 1;
    CollectInput(RESET:=TRUE);
  END_IF;
END_PROGRAM

CONFIGURATION Config0
  RESOURCE Res0 ON PLC
    TASK task0(INTERVAL := T#20ms,PRIORITY := 0);
    PROGRAM instance0 WITH task0 : Boiler;
  END_RESOURCE
END_CONFIGURATION

(* ---- RND-EXPR_alias-snake-bodge.st ---- *)
(*
This code implements a randomly grown symbolic expression:

IN38 | IN6

*)

FUNCTION_BLOCK F_CollectInput
  VAR_IN_OUT
      Data : ARRAY[1..50] OF BOOL;
  END_VAR
  VAR_INPUT
      TICK  : BOOL := 0;
      IN1   : BOOL := 0;
      IN2   : BOOL := 0;
      IN3   : BOOL := 0;
      IN4   : BOOL := 0;
      IN5   : BOOL := 0;
      RESET : BOOL := FALSE;
  END_VAR
  VAR_OUTPUT
      Finished : BOOL;
  END_VAR
  VAR
      j    : USINT := 1;
      tock : BOOL  := 0;
  END_VAR
  IF NOT RESET AND tock = NOT TICK THEN
      Data[j]   := IN1;
      Data[j+1] := IN2;
      Data[j+2] := IN3;
      Data[j+3] := IN4;
      Data[j+4] := IN5;
      j := j + 5;
      tock := TICK;
  ELSE
      j := 1;
      tock := 0;
  END_IF;
  Finished := (j > 50);
END_FUNCTION_BLOCK

PROGRAM Boiler
  VAR
    Data  : ARRAY[1..50] OF BOOL;
    Ready : BOOL;
    CollectInput : F_CollectInput;
  END_VAR
  VAR
    TICK     AT %IX1.0 : BOOL;
    IN1      AT %IX0.3 : BOOL;
    IN2      AT %IX0.4 : BOOL;
    IN3      AT %IX0.5 : BOOL;
    IN4      AT %IX0.6 : BOOL;
    IN5      AT %IX0.7 : BOOL;
    OutReady AT %QX0.0 : BOOL := FALSE;
    FeedNext AT %QX0.1 : BOOL := FALSE;
    Out      AT %QX0.2 : BOOL;
  END_VAR
  CollectInput(TICK:=TICK, IN1:=IN1, IN2:=IN2, IN3:=IN3, IN4:=IN4, IN5:=IN5);
  Ready := CollectInput.Finished;
  FeedNext := 1;
  IF Ready THEN
    Out := (Data[38] OR Data[6]);
    OutReady := 1;
    CollectInput(RESET:=TRUE);
  END_IF;
END_PROGRAM

CONFIGURATION Config0
  RESOURCE Res0 ON PLC
    TASK task0(INTERVAL := T#20ms,PRIORITY := 0);
    PROGRAM instance0 WITH task0 : Boiler;
  END_RESOURCE
END_CONFIGURATION
